METHOD PRIVATE PublishHmi
// Единый снимок состояния для внешней визуализации.
GVL_HMI.udiPlcHeartbeat := GVL_HMI.udiPlcHeartbeat + 1;
GVL_HMI.xHmiConnectionAlive := xHmiConnectionAlive;
GVL_HMI.xManualRecoveryActive := xManualRecoveryActive;
GVL_HMI.xGlobalError := GVL_CELL_CONTROL.xGlobalError;
GVL_HMI.xCellManual := GVL_CELL_CONTROL.xManual;
// Отказ тоже потребляет транзакцию: она не исполнится позже сама собой.
GVL_HMI.udiCellModeAckSeq := udiCellModeCommandSnapshot;
GVL_HMI.xErrorSimulationEnabled := GVL_CELL_SETTINGS.xErrorSimulationEnabled;
GVL_HMI.stSafetyFaultStatus := CELL_SAFETY.FaultStatus;
GVL_HMI.xSimulationAccelerationActive := GVL_CELL_SETTINGS.xSimulationAccelerationActive;
GVL_HMI.xSimulationAccelerationChangeAllowed := GVL_CELL_SETTINGS.xSimulationAccelerationChangeAllowed;
GVL_HMI.uiSimulationTimeFactorApplied := GVL_CELL_SETTINGS.uiSimulationTimeFactorApplied;
GVL_HMI.xSimulationAccelerationPending := GVL_CELL_SETTINGS.xSimulationAccelerationPending;
GVL_HMI.xSimulationAccelerationBusy := GVL_CELL_SETTINGS.xSimulationAccelerationBusy;
GVL_HMI.xSimulationAccelerationError := GVL_CELL_SETTINGS.xSimulationAccelerationError;
GVL_HMI.udiSimulationAccelerationErrorId := GVL_CELL_SETTINGS.udiSimulationAccelerationErrorId;
GVL_HMI.lrSafetyHomeX := GVL_POINT.Points[E_POINT_NAME.HOME_SAFETY].X;
GVL_HMI.lrSafetyHomeY := GVL_POINT.Points[E_POINT_NAME.HOME_SAFETY].Y;
GVL_HMI.lrSafetyHomeZ := GVL_POINT.Points[E_POINT_NAME.HOME_SAFETY].Z;
GVL_HMI.lrSafetyHomeSpeedFactor := GVL_POINT.Points[E_POINT_NAME.HOME_SAFETY].SpeedFactor;
GVL_HMI.lrSafetyHomeToleranceX := GVL_CELL_SETTINGS.lrSafetyHomeToleranceX;
GVL_HMI.lrSafetyHomeToleranceY := GVL_CELL_SETTINGS.lrSafetyHomeToleranceY;
GVL_HMI.lrSafetyHomeToleranceZ := GVL_CELL_SETTINGS.lrSafetyHomeToleranceZ;
GVL_HMI.rRobotAccelerationPercent := GVL_CELL_SETTINGS.rRobotAccelerationPercent;
GVL_HMI.rRobotDecelerationPercent := GVL_CELL_SETTINGS.rRobotDecelerationPercent;
GVL_HMI.rRobotJerkPercent := GVL_CELL_SETTINGS.rRobotJerkPercent;
GVL_HMI.lrRobotHaltDeceleration := GVL_CELL_SETTINGS.lrRobotHaltDeceleration;
GVL_HMI.lrRobotHaltJerk := GVL_CELL_SETTINGS.lrRobotHaltJerk;
GVL_HMI.stCellMachineTimeouts := GVL_CELL_SETTINGS.stMachineTimeouts;
GVL_HMI.stCellAxisTimeouts := GVL_CELL_SETTINGS.stAxisTimeouts;
GVL_HMI.stCellAxisGroupTimeouts := GVL_CELL_SETTINGS.stAxisGroupTimeouts;
GVL_HMI.tPointCheckStartTimeout := GVL_CELL_SETTINGS.tPointCheckStartTimeout;
GVL_HMI.tSimulationDynamicsTimeout := GVL_CELL_SETTINGS.tSimulationDynamicsTimeout;
GVL_HMI.tHmiWatchdogTimeout := GVL_CELL_SETTINGS.tHmiWatchdogTimeout;
GVL_HMI.tMobileMotionWatchdogTimeout := GVL_CELL_SETTINGS.tMobileMotionWatchdogTimeout;
GVL_HMI.tPointCheckWatchdogTimeout := GVL_CELL_SETTINGS.tPointCheckWatchdogTimeout;
GVL_HMI.tHmiCommandFreshnessTimeout := GVL_CELL_SETTINGS.tHmiCommandFreshnessTimeout;
GVL_HMI.tAlarmHornDuration := GVL_CELL_SETTINGS.tAlarmHornDuration;
GVL_HMI.tInputFilterRise := GVL_CELL_SETTINGS.tInputFilterRise;
GVL_HMI.tInputFilterFall := GVL_CELL_SETTINGS.tInputFilterFall;
GVL_HMI.xIoFilterSettingsChangeAllowed := GVL_CELL_SETTINGS.xIoFilterSettingsChangeAllowed;
GVL_HMI.xPhysicalIoActive := GVL_PHYSICAL_IO.xNormalActive
	AND (GVL_CELL_SETTINGS.eTestEnvironment = E_CELL_TEST_ENVIRONMENT.NORMAL);
GVL_HMI.xPhysicalIoMappingVerified := GVL_PHYSICAL_IO.xMappingVerified;
GVL_HMI.xCellSettingsChangeAllowed := GVL_CELL_SETTINGS.xCellSettingsChangeAllowed;
GVL_HMI.rPointCheckSpeedPercent := GVL_CELL_SETTINGS.rPointCheckSpeedPercent;
GVL_HMI.xPointCheckActive := xPointCheckActive;
IF xPointCheckActive THEN
	GVL_HMI.rPointCheckAppliedSpeedPercent := rPointCheckLatchedSpeed;
ELSE
	GVL_HMI.rPointCheckAppliedSpeedPercent := GVL_CELL_SETTINGS.rPointCheckSpeedPercent;
END_IF;
GVL_HMI.xPointTableReady := xPointTableReady;
GVL_HMI.astPointEditorPoints[1] := GVL_POINT.Points[E_POINT_NAME.MACHINE_1_ABOVE];
GVL_HMI.astPointEditorPoints[2] := GVL_POINT.Points[E_POINT_NAME.MACHINE_1_CHUCK_APROACH];
GVL_HMI.astPointEditorPoints[3] := GVL_POINT.Points[E_POINT_NAME.MACHINE_1_CHUCK_POSITION];
GVL_HMI.astPointEditorPoints[4] := GVL_POINT.Points[E_POINT_NAME.MACHINE_2_ABOVE];
GVL_HMI.astPointEditorPoints[5] := GVL_POINT.Points[E_POINT_NAME.MACHINE_2_CHUCK_APROACH];
GVL_HMI.astPointEditorPoints[6] := GVL_POINT.Points[E_POINT_NAME.MACHINE_2_CHUCK_POSITION];
GVL_HMI.astPointEditorPoints[7] := GVL_POINT.Points[E_POINT_NAME.MACHINE_3_ABOVE];
GVL_HMI.astPointEditorPoints[8] := GVL_POINT.Points[E_POINT_NAME.MACHINE_3_CHUCK_APROACH];
GVL_HMI.astPointEditorPoints[9] := GVL_POINT.Points[E_POINT_NAME.MACHINE_3_CHUCK_POSITION];
GVL_HMI.astPointEditorPoints[10] := GVL_POINT.Points[E_POINT_NAME.HOME_SAFETY];
GVL_HMI.astPointEditorPoints[11] := GVL_POINT.Points[E_POINT_NAME.MAGAZINE_1_DETAIL];
GVL_HMI.astPointEditorPoints[12] := GVL_POINT.Points[E_POINT_NAME.MAGAZINE_2_DETAIL];
GVL_HMI.astPointEditorPoints[13] := GVL_POINT.Points[E_POINT_NAME.GEOMETRY_1_PLACE];
GVL_HMI.astPointEditorPoints[14] := GVL_POINT.Points[E_POINT_NAME.GEOMETRY_2_PLACE];
GVL_HMI.auiPointEditorPointId[1] := TO_UINT(E_POINT_NAME.MACHINE_1_ABOVE);
GVL_HMI.auiPointEditorPointId[2] := TO_UINT(E_POINT_NAME.MACHINE_1_CHUCK_APROACH);
GVL_HMI.auiPointEditorPointId[3] := TO_UINT(E_POINT_NAME.MACHINE_1_CHUCK_POSITION);
GVL_HMI.auiPointEditorPointId[4] := TO_UINT(E_POINT_NAME.MACHINE_2_ABOVE);
GVL_HMI.auiPointEditorPointId[5] := TO_UINT(E_POINT_NAME.MACHINE_2_CHUCK_APROACH);
GVL_HMI.auiPointEditorPointId[6] := TO_UINT(E_POINT_NAME.MACHINE_2_CHUCK_POSITION);
GVL_HMI.auiPointEditorPointId[7] := TO_UINT(E_POINT_NAME.MACHINE_3_ABOVE);
GVL_HMI.auiPointEditorPointId[8] := TO_UINT(E_POINT_NAME.MACHINE_3_CHUCK_APROACH);
GVL_HMI.auiPointEditorPointId[9] := TO_UINT(E_POINT_NAME.MACHINE_3_CHUCK_POSITION);
GVL_HMI.auiPointEditorPointId[10] := TO_UINT(E_POINT_NAME.HOME_SAFETY);
GVL_HMI.auiPointEditorPointId[11] := TO_UINT(E_POINT_NAME.MAGAZINE_1_DETAIL);
GVL_HMI.auiPointEditorPointId[12] := TO_UINT(E_POINT_NAME.MAGAZINE_2_DETAIL);
GVL_HMI.auiPointEditorPointId[13] := TO_UINT(E_POINT_NAME.GEOMETRY_1_PLACE);
GVL_HMI.auiPointEditorPointId[14] := TO_UINT(E_POINT_NAME.GEOMETRY_2_PLACE);
GVL_HMI.xModbusMode := GVL_ROBOT_MODBUS.xModeActive;
GVL_HMI.xRobotModeChangeAllowed := GVL_ROBOT_MODBUS.xRobotModeChangeAllowed;
GVL_HMI.xModbusSettingsChangeAllowed := GVL_ROBOT_MODBUS.xSettingsChangeAllowed;
GVL_HMI.stRobotModbusStatus := GVL_ROBOT_MODBUS.Status;
uiMagazine := GVL_CELL_MANAGER.Status.uiActiveMagazine;
IF (uiMagazine < UINT#1) OR (uiMagazine > UINT#2) THEN
	uiMagazine := UINT#1;
END_IF;
GVL_HMI.stTestObservability.udiAppliedScenarioSeq := GVL_HMI.udiTestScenarioAckSeq;
GVL_HMI.stTestObservability.uiCellState := TO_UINT(GVL_CELL_MANAGER.Diag.eState);
GVL_HMI.stTestObservability.uiRobotState := TO_UINT(GVL_ROBOT.Diag.eState);
GVL_HMI.stTestObservability.uiRobotAction := TO_UINT(GVL_ROBOT.Diag.eActiveAction);
GVL_HMI.stTestObservability.uiRobotPoint := TO_UINT(GVL_ROBOT.Diag.eActivePoint);
GVL_HMI.stTestObservability.uiActiveMagazine := GVL_CELL_MANAGER.Status.uiActiveMagazine;
GVL_HMI.stTestObservability.uiMagazineState := TO_UINT(GVL_MAGAZINE.astDiag[uiMagazine].eState);
GVL_HMI.stTestObservability.uiMagazineOperation := TO_UINT(GVL_MAGAZINE.astStatus[uiMagazine].eActualOperation);
GVL_HMI.stTestObservability.uiTakeSlot := SINT_TO_UINT(GVL_MAGAZINE.astStatus[uiMagazine].iSelectedBlank);
GVL_HMI.stTestObservability.uiPutSlot := SINT_TO_UINT(GVL_MAGAZINE.astStatus[uiMagazine].iSelectedFreeSlot);
GVL_HMI.stTestObservability.uiSelectedMachine := GVL_CELL_MANAGER.Status.uiSelectedMachine;
GVL_HMI.stTestObservability.uiSelectedType := GVL_MULTI_TYPE.CycleStatus.uiSelectedType;
GVL_HMI.stTestObservability.uiErrorSource := UINT#0;
GVL_HMI.stTestObservability.dwErrorCode := DWORD#0;
FOR uiMachine := 1 TO 3 DO
	GVL_HMI.stTestObservability.auiMachineState[uiMachine] := TO_UINT(GVL_MACHINE.Diag[uiMachine].eState);
	GVL_HMI.stTestObservability.auiMachineOperation[uiMachine] := TO_UINT(GVL_MACHINE.Diag[uiMachine].eActualOperation);
END_FOR;
IF GVL_ROBOT.Error.dwErrorActive <> DWORD#0 THEN
	GVL_HMI.stTestObservability.uiErrorSource := UINT#2;
	GVL_HMI.stTestObservability.dwErrorCode := GVL_ROBOT.Error.dwErrorActive;
ELSIF GVL_MAGAZINE.astError[1].dwErrorActive <> DWORD#0 THEN
	GVL_HMI.stTestObservability.uiErrorSource := UINT#3;
GVL_HMI.stTestObservability.dwErrorCode := GVL_MAGAZINE.astError[1].dwErrorActive;
ELSIF GVL_MAGAZINE.astError[2].dwErrorActive <> DWORD#0 THEN
	GVL_HMI.stTestObservability.uiErrorSource := UINT#7;
	GVL_HMI.stTestObservability.dwErrorCode := GVL_MAGAZINE.astError[2].dwErrorActive;
ELSIF GVL_CELL_MANAGER.Error.dwErrorActive <> DWORD#0 THEN
	GVL_HMI.stTestObservability.uiErrorSource := UINT#1;
	GVL_HMI.stTestObservability.dwErrorCode := GVL_CELL_MANAGER.Error.dwErrorActive;
ELSE
	FOR uiMachine := 1 TO 3 DO
		IF GVL_MACHINE.Error[uiMachine].dwErrorActive <> DWORD#0 THEN
			GVL_HMI.stTestObservability.uiErrorSource := uiMachine + UINT#3;
			GVL_HMI.stTestObservability.dwErrorCode := GVL_MACHINE.Error[uiMachine].dwErrorActive;
		END_IF;
	END_FOR;
END_IF;
FOR uiMachine := 1 TO 9 DO
	GVL_HMI.auiRobotModbusWriteRegisters[uiMachine] :=
		GVL_ROBOT_MODBUS.auiWriteRegisters[uiMachine - 1];
END_FOR;
FOR uiMachine := 1 TO 17 DO
	GVL_HMI.auiRobotModbusReadRegisters[uiMachine] :=
		GVL_ROBOT_MODBUS.auiReadRegisters[uiMachine - 1];
END_FOR;
GVL_HMI.xSimAxisGroupErrorAllowed := GVL_AXIS_GROUP.AxisGroup.Status.xSimErrorAllowed;
GVL_HMI.astAxisFaultStatus[1] := AXIS_X.FaultStatus;
GVL_HMI.astAxisFaultStatus[2] := AXIS_Y.FaultStatus;
GVL_HMI.astAxisFaultStatus[3] := AXIS_Z.FaultStatus;
GVL_HMI.stAxisGroupFaultStatus := GROUP_XYZ.FaultStatus;
GVL_HMI.stGripperFaultStatus := ROBOT.FaultStatus.stGripper;
GVL_HMI.stRobotFaultStatus := ROBOT.FaultStatus.stRobot;
GVL_HMI.stCellFaultStatus := CELL_MANAGER.FaultStatus;
GVL_HMI.stPointFaultStatus := ROBOT.FaultStatus.stPoint;
GVL_HMI.stMagazineFaultStatus := fbMagazine1.FaultStatus;
GVL_HMI.astMagazineFaultStatus[1] := fbMagazine1.FaultStatus;
GVL_HMI.astMagazineFaultStatus[2] := fbMagazine2.FaultStatus;
GVL_HMI.rLoadCNC_1 := GVL_STATISTIC.stStatistic.stMachineStat.rLoadCNC_1;
GVL_HMI.rLoadCNC_2 := GVL_STATISTIC.stStatistic.stMachineStat.rLoadCNC_2;
GVL_HMI.rLoadCNC_3 := GVL_STATISTIC.stStatistic.stMachineStat.rLoadCNC_3;
GVL_HMI.rRobot := GVL_STATISTIC.stStatistic.stRobotStat.rRobot;

GVL_HMI.stCellStatus := GVL_CELL_MANAGER.Status;
GVL_HMI.stCellStatus.xResetAllowed := xAlarmResetAllowed;
GVL_HMI.stCellDiag := GVL_CELL_MANAGER.Diag;
GVL_HMI.stCellError := GVL_CELL_MANAGER.Error;
GVL_HMI.stCellSafetyStatus := CELL_SAFETY.Status;
GVL_HMI.stCellSafetyDiag := CELL_SAFETY.Diag;
GVL_HMI.stCellSafetyError := CELL_SAFETY.Error;
GVL_HMI.astButtonStationIoStatus := CELL_SAFETY.astButtonStationIoStatus;
GVL_HMI.stFrontControlCabinetIoStatus := CELL_SAFETY.stFrontControlCabinetIoStatus;
GVL_HMI.xSignalTowerRed := GVL_CELL_SAFETY_IO.xSignalTowerRedOutput;
GVL_HMI.xSignalTowerAmber := GVL_CELL_SAFETY_IO.xSignalTowerAmberOutput;
GVL_HMI.xSignalTowerGreen := GVL_CELL_SAFETY_IO.xSignalTowerGreenOutput;
GVL_HMI.stRearControlCabinetIoStatus := CELL_SAFETY.stRearControlCabinetIoStatus;
GVL_HMI.stMpgIoStatus := CELL_SAFETY.stMpgIoStatus;
GVL_HMI.astEnclosureDoorStatus := CELL_SAFETY.astEnclosureDoorStatus;
GVL_HMI.stMultiType.Config := GVL_MULTI_TYPE.Config;
GVL_HMI.stMultiType.ConfigStatus := GVL_MULTI_TYPE.ConfigStatus;
GVL_HMI.stMultiType.CycleStatus := GVL_MULTI_TYPE.CycleStatus;

GVL_HMI.stRobotStatus := GVL_ROBOT.Status;
GVL_HMI.stRobotDiag := GVL_ROBOT.Diag;
GVL_HMI.stRobotError := GVL_ROBOT.Error;
GVL_HMI.stGripperDiag := GVL_ROBOT.GripperDiag;
GVL_HMI.stGripperError := GVL_ROBOT.GripperError;
GVL_HMI.stAxisGroupStatus := GVL_AXIS_GROUP.AxisGroup.Status;
GVL_HMI.stAxisGroupDiag := GVL_AXIS_GROUP.AxisGroup.Diag;
GVL_HMI.stAxisGroupError := GVL_AXIS_GROUP.AxisGroup.Error;
GVL_HMI.stMotionManagerStatus := GVL_MOTION_MANAGER.stMotionManager.Status;
GVL_HMI.stMotionManagerDiag := GVL_MOTION_MANAGER.stMotionManager.Diag;
GVL_HMI.stMotionManagerError := GVL_MOTION_MANAGER.stMotionManager.Error;
GVL_HMI.stPointManagerStatus := GVL_POINT_MANAGER.PointManager.Status;
GVL_HMI.stPointManagerDiag := GVL_POINT_MANAGER.PointManager.Diag;
GVL_HMI.stPointManagerError := GVL_POINT_MANAGER.PointManager.Error;

FOR uiMachine := 1 TO 3 DO
	GVL_HMI.astAxisStatus[uiMachine] := GVL_AXIS.arrAxis[uiMachine].Status;
	GVL_HMI.astAxisDiag[uiMachine] := GVL_AXIS.arrAxis[uiMachine].Diag;
	GVL_HMI.astAxisError[uiMachine] := GVL_AXIS.arrAxis[uiMachine].Error;
END_FOR;

GVL_HMI.stMagazineStatus := GVL_MAGAZINE.astStatus[1];
GVL_HMI.stMagazineDiag := GVL_MAGAZINE.astDiag[1];
GVL_HMI.stMagazineError := GVL_MAGAZINE.astError[1];
FOR uiMagazine := UINT#1 TO UINT#2 DO
	GVL_HMI.astMagazineStatus[uiMagazine] := GVL_MAGAZINE.astStatus[uiMagazine];
	GVL_HMI.astMagazineDiag[uiMagazine] := GVL_MAGAZINE.astDiag[uiMagazine];
	GVL_HMI.astMagazineError[uiMagazine] := GVL_MAGAZINE.astError[uiMagazine];
	GVL_HMI.astMagazineInventory[uiMagazine] := GVL_DETAIL.astMagazine[uiMagazine];
END_FOR;
GVL_HMI.stAlarmStatus := GVL_ALARM.Status;
GVL_HMI.astAlarmEvent := GVL_ALARM.Events;

FOR uiMachine := 1 TO 3 DO
	GVL_HMI.astMachineStatus[uiMachine] := GVL_MACHINE.Status[uiMachine];
	GVL_HMI.astMachineDiag[uiMachine] := GVL_MACHINE.Diag[uiMachine];
	GVL_HMI.astMachineError[uiMachine] := GVL_MACHINE.Error[uiMachine];
	CASE uiMachine OF
		1:
			GVL_HMI.astMachineFaultStatus[uiMachine] := MACHINE_1_FAULT.Status;
			GVL_HMI.astMachineFaultStatus[uiMachine].xResetAllowed :=
				MACHINE_1_SIM.Diag.xResetAllowed OR GVL_MACHINE.Status[uiMachine].xResetAllowed;
		2:
			GVL_HMI.astMachineFaultStatus[uiMachine] := MACHINE_2_FAULT.Status;
			GVL_HMI.astMachineFaultStatus[uiMachine].xResetAllowed :=
				MACHINE_2_SIM.Diag.xResetAllowed OR GVL_MACHINE.Status[uiMachine].xResetAllowed;
		3:
			GVL_HMI.astMachineFaultStatus[uiMachine] := MACHINE_3_FAULT.Status;
			GVL_HMI.astMachineFaultStatus[uiMachine].xResetAllowed :=
				MACHINE_3_SIM.Diag.xResetAllowed OR GVL_MACHINE.Status[uiMachine].xResetAllowed;
	END_CASE;
END_FOR;

GVL_HMI.astMachineIoStatus[1] := MACHINE_1_FAULT.MachineStatus;
GVL_HMI.astMachineIoStatus[2] := MACHINE_2_FAULT.MachineStatus;
GVL_HMI.astMachineIoStatus[3] := MACHINE_3_FAULT.MachineStatus;
GVL_HMI.astMachineRawIoStatus[1] := MACHINE_1_SIM.Status;
GVL_HMI.astMachineRawIoStatus[2] := MACHINE_2_SIM.Status;
GVL_HMI.astMachineRawIoStatus[3] := MACHINE_3_SIM.Status;
GVL_HMI.astMachineTimeouts[1] := MACHINE_1_FAULT.Timeouts;
GVL_HMI.astMachineTimeouts[2] := MACHINE_2_FAULT.Timeouts;
GVL_HMI.astMachineTimeouts[3] := MACHINE_3_FAULT.Timeouts;
GVL_HMI.astMachineSimDiag[1] := MACHINE_1_SIM.Diag;
GVL_HMI.astMachineSimDiag[2] := MACHINE_2_SIM.Diag;
GVL_HMI.astMachineSimDiag[3] := MACHINE_3_SIM.Diag;
GVL_HMI.astMachineSimError[1] := MACHINE_1_SIM.Error;
GVL_HMI.astMachineSimError[2] := MACHINE_2_SIM.Error;
GVL_HMI.astMachineSimError[3] := MACHINE_3_SIM.Error;

FOR iDetail := 1 TO GVL_CELL_SETTINGS.NumberDetail DO
	GVL_HMI.astMagazineSlot[iDetail] := GVL_DETAIL.astMagazine[1].aSlots[iDetail];
END_FOR;

// Ack only the snapshot actually dispatched through all consumers this scan.
FOR uiHmiCommandIndex := UINT#1 TO UINT#121 DO
	IF axHmiCommandConsumed[uiHmiCommandIndex] THEN
		GVL_HMI.audiHmiCommandAckSeq[uiHmiCommandIndex] := audiHmiCommandSnapshot[uiHmiCommandIndex];
	END_IF;
END_FOR;
GVL_HMI.udiCellSettingAckSeq := udiCellSettingSnapshot;

GVL_HMI.uiMagazineMode := GVL_TWO_PALLET.uiMode;
GVL_HMI.xMagazineModeAllowed := GVL_TWO_PALLET.xModeChangeAllowed;
GVL_HMI.astTwinStatus := GVL_TWO_PALLET.astStatus;
GVL_HMI.astTwinConfig := GVL_TWO_PALLET.astActiveConfig;
GVL_HMI.astTwinStore := GVL_TWO_PALLET.astStore;
END_METHOD

METHOD PRIVATE IsHmiCommandFresh : BOOL
VAR_INPUT
	udiIssuedAtMs : UDINT;
END_VAR
VAR
	uliAgeMs : ULINT;
END_VAR
// Explicit modulo-2^32 age: TIME() rolls over after about 49 days.
IF udiHmiCommandNowMs >= udiIssuedAtMs THEN
	uliAgeMs := UDINT_TO_ULINT(udiHmiCommandNowMs) - UDINT_TO_ULINT(udiIssuedAtMs);
ELSE
	uliAgeMs := ULINT#4294967296 + UDINT_TO_ULINT(udiHmiCommandNowMs) - UDINT_TO_ULINT(udiIssuedAtMs);
END_IF;
IsHmiCommandFresh := uliAgeMs <= UDINT_TO_ULINT(
	TIME_TO_UDINT(GVL_CELL_SETTINGS.tHmiCommandFreshnessTimeout)
);
END_METHOD

METHOD PRIVATE WritePhysicalOutputs
// Единственная страница назначения выходов. Выполняется после всех владельцев команд.
// Не публикуем команды симулятора на железо при смене среды в текущем скане.
xPhysicalOutputEnable := GVL_PHYSICAL_IO.xNormalActive
	AND (GVL_CELL_SETTINGS.eTestEnvironment = E_CELL_TEST_ENVIRONMENT.NORMAL);
IF xPhysicalOutputEnable THEN
	FOR uiMachine := 1 TO 3 DO
		IF GVL_MACHINE.Command[uiMachine].stIo.xCloseDoor
		AND NOT GVL_MACHINE.Command[uiMachine].stIo.xOpenDoor THEN
			GVL_PHYSICAL_IO.axMachineHatchClose[uiMachine] := TRUE;
		ELSIF GVL_MACHINE.Command[uiMachine].stIo.xOpenDoor
		AND NOT GVL_MACHINE.Command[uiMachine].stIo.xCloseDoor THEN
			GVL_PHYSICAL_IO.axMachineHatchClose[uiMachine] := FALSE;
		ELSIF NOT xPhysicalOutputWasEnabled THEN
			GVL_PHYSICAL_IO.axMachineHatchClose[uiMachine] := GVL_MACHINE.astPhysicalInput[uiMachine].xDoorClosed;
		END_IF;
	END_FOR;
	IF NOT GVL_HMI.xModbusMode AND GVL_PHYSICAL_IO.stGripperCommand.xExecute THEN
		CASE GVL_PHYSICAL_IO.stGripperCommand.eAction OF
			E_ROBOT_ACTION.UNCLAMP_1: axIoGripperBase[1] := TRUE;
			E_ROBOT_ACTION.CLAMP_1: axIoGripperBase[1] := FALSE;
			E_ROBOT_ACTION.UNCLAMP_2: axIoGripperBase[2] := TRUE;
			E_ROBOT_ACTION.CLAMP_2: axIoGripperBase[2] := FALSE;
			E_ROBOT_ACTION.ROTATE_TO_BLANK: axIoGripperBase[3] := FALSE;
			E_ROBOT_ACTION.ROTATE_TO_DETAIL: axIoGripperBase[3] := TRUE;
		END_CASE;
	END_IF;
END_IF;
// Внешний SC-500 остаётся единственным владельцем захватов в Modbus.
IF NOT xPhysicalOutputEnable OR GVL_HMI.xModbusMode THEN
	axIoGripperBase[1] := FALSE;
	axIoGripperBase[2] := FALSE;
	axIoGripperBase[3] := FALSE;
END_IF;
GVL_PHYSICAL_IO.xDoGripper1Open := axIoGripperBase[1];
GVL_PHYSICAL_IO.xDoGripper2Open := axIoGripperBase[2];
GVL_PHYSICAL_IO.xDoRotateToDetail := axIoGripperBase[3];

GVL_PHYSICAL_IO.xDoMachine1HatchClosed := xPhysicalOutputEnable AND GVL_PHYSICAL_IO.axMachineHatchClose[1];
GVL_PHYSICAL_IO.xDoMachine1HatchUnLock := xPhysicalOutputEnable AND GVL_MACHINE.Command[1].stIo.xHatchUnLock;
GVL_PHYSICAL_IO.xDoMachine1ClampChuck := xPhysicalOutputEnable AND GVL_MACHINE.Command[1].stIo.xClampChuck AND NOT GVL_MACHINE.Command[1].stIo.xUnclampChuck;
GVL_PHYSICAL_IO.xDoMachine1UnclampChuck := xPhysicalOutputEnable AND GVL_MACHINE.Command[1].stIo.xUnclampChuck AND NOT GVL_MACHINE.Command[1].stIo.xClampChuck;
GVL_PHYSICAL_IO.xDoMachine1StartCycle := xPhysicalOutputEnable AND GVL_MACHINE.Command[1].stIo.xStartCycle;
GVL_PHYSICAL_IO.xDoMachine2HatchClosed := xPhysicalOutputEnable AND GVL_PHYSICAL_IO.axMachineHatchClose[2];
GVL_PHYSICAL_IO.xDoMachine2HatchUnLock := xPhysicalOutputEnable AND GVL_MACHINE.Command[2].stIo.xHatchUnLock;
GVL_PHYSICAL_IO.xDoMachine2ClampChuck := xPhysicalOutputEnable AND GVL_MACHINE.Command[2].stIo.xClampChuck AND NOT GVL_MACHINE.Command[2].stIo.xUnclampChuck;
GVL_PHYSICAL_IO.xDoMachine2UnclampChuck := xPhysicalOutputEnable AND GVL_MACHINE.Command[2].stIo.xUnclampChuck AND NOT GVL_MACHINE.Command[2].stIo.xClampChuck;
GVL_PHYSICAL_IO.xDoMachine2StartCycle := xPhysicalOutputEnable AND GVL_MACHINE.Command[2].stIo.xStartCycle;
GVL_PHYSICAL_IO.xDoMachine3HatchClosed := xPhysicalOutputEnable AND GVL_PHYSICAL_IO.axMachineHatchClose[3];
GVL_PHYSICAL_IO.xDoMachine3HatchUnLock := xPhysicalOutputEnable AND GVL_MACHINE.Command[3].stIo.xHatchUnLock;
GVL_PHYSICAL_IO.xDoMachine3ClampChuck := xPhysicalOutputEnable AND GVL_MACHINE.Command[3].stIo.xClampChuck AND NOT GVL_MACHINE.Command[3].stIo.xUnclampChuck;
GVL_PHYSICAL_IO.xDoMachine3UnclampChuck := xPhysicalOutputEnable AND GVL_MACHINE.Command[3].stIo.xUnclampChuck AND NOT GVL_MACHINE.Command[3].stIo.xClampChuck;
GVL_PHYSICAL_IO.xDoMachine3StartCycle := xPhysicalOutputEnable AND GVL_MACHINE.Command[3].stIo.xStartCycle;
GVL_PHYSICAL_IO.xDoDoor1Unlock := xPhysicalOutputEnable AND GVL_CELL_SAFETY_IO.axDoorUnlockOutput[1];
GVL_PHYSICAL_IO.xDoDoor2Unlock := xPhysicalOutputEnable AND GVL_CELL_SAFETY_IO.axDoorUnlockOutput[2];
GVL_PHYSICAL_IO.xDoDoor3Unlock := xPhysicalOutputEnable AND GVL_CELL_SAFETY_IO.axDoorUnlockOutput[3];
GVL_PHYSICAL_IO.xDoDoor4Unlock := xPhysicalOutputEnable AND GVL_CELL_SAFETY_IO.axDoorUnlockOutput[4];
GVL_PHYSICAL_IO.xDoSafetyRelayReset := xPhysicalOutputEnable AND GVL_CELL_SAFETY_IO.xSafetyRelayResetOutput;
GVL_PHYSICAL_IO.xDoSignalTowerGreenOutput := xPhysicalOutputEnable AND GVL_CELL_SAFETY_IO.xSignalTowerGreenOutput;
GVL_PHYSICAL_IO.xDoSignalTowerAmberOutput := xPhysicalOutputEnable AND GVL_CELL_SAFETY_IO.xSignalTowerAmberOutput;
GVL_PHYSICAL_IO.xDoSignalTowerRedOutput := xPhysicalOutputEnable AND GVL_CELL_SAFETY_IO.xSignalTowerRedOutput;
GVL_PHYSICAL_IO.xDoDoor1ButtonLamp := xPhysicalOutputEnable AND GVL_CELL_SAFETY_IO.axDoorButtonLampOutput[1];
GVL_PHYSICAL_IO.xDoDoor2ButtonLamp := xPhysicalOutputEnable AND GVL_CELL_SAFETY_IO.axDoorButtonLampOutput[2];
GVL_PHYSICAL_IO.xDoDoor3ButtonLamp := xPhysicalOutputEnable AND GVL_CELL_SAFETY_IO.axDoorButtonLampOutput[3];
GVL_PHYSICAL_IO.xDoDoor4ButtonLamp := xPhysicalOutputEnable AND GVL_CELL_SAFETY_IO.axDoorButtonLampOutput[4];
GVL_PHYSICAL_IO.xDoMagazine1LockIn := xPhysicalOutputEnable AND (GVL_TWO_PALLET.uiMode = UINT#1) AND GVL_TWO_PALLET.astOutput[1].xLockIn AND NOT GVL_TWO_PALLET.astOutput[1].xLockOut;
GVL_PHYSICAL_IO.xDoMagazine1LockOut := xPhysicalOutputEnable AND (GVL_TWO_PALLET.uiMode = UINT#1) AND GVL_TWO_PALLET.astOutput[1].xLockOut AND NOT GVL_TWO_PALLET.astOutput[1].xLockIn;
GVL_PHYSICAL_IO.xDoMagazine1StopIn := xPhysicalOutputEnable AND (GVL_TWO_PALLET.uiMode = UINT#1) AND GVL_TWO_PALLET.astOutput[1].xStopIn AND NOT GVL_TWO_PALLET.astOutput[1].xStopOut;
GVL_PHYSICAL_IO.xDoMagazine1StopOut := xPhysicalOutputEnable AND (GVL_TWO_PALLET.uiMode = UINT#1) AND GVL_TWO_PALLET.astOutput[1].xStopOut AND NOT GVL_TWO_PALLET.astOutput[1].xStopIn;
GVL_PHYSICAL_IO.xDoMagazine1LiftUp := xPhysicalOutputEnable AND (GVL_TWO_PALLET.uiMode = UINT#1) AND GVL_TWO_PALLET.astOutput[1].xLiftUp AND NOT GVL_TWO_PALLET.astOutput[1].xLiftDown;
GVL_PHYSICAL_IO.xDoMagazine1LiftDown := xPhysicalOutputEnable AND (GVL_TWO_PALLET.uiMode = UINT#1) AND GVL_TWO_PALLET.astOutput[1].xLiftDown AND NOT GVL_TWO_PALLET.astOutput[1].xLiftUp;
GVL_PHYSICAL_IO.xDoMagazine2LockIn := xPhysicalOutputEnable AND (GVL_TWO_PALLET.uiMode = UINT#1) AND GVL_TWO_PALLET.astOutput[2].xLockIn AND NOT GVL_TWO_PALLET.astOutput[2].xLockOut;
GVL_PHYSICAL_IO.xDoMagazine2LockOut := xPhysicalOutputEnable AND (GVL_TWO_PALLET.uiMode = UINT#1) AND GVL_TWO_PALLET.astOutput[2].xLockOut AND NOT GVL_TWO_PALLET.astOutput[2].xLockIn;
GVL_PHYSICAL_IO.xDoMagazine2StopIn := xPhysicalOutputEnable AND (GVL_TWO_PALLET.uiMode = UINT#1) AND GVL_TWO_PALLET.astOutput[2].xStopIn AND NOT GVL_TWO_PALLET.astOutput[2].xStopOut;
GVL_PHYSICAL_IO.xDoMagazine2StopOut := xPhysicalOutputEnable AND (GVL_TWO_PALLET.uiMode = UINT#1) AND GVL_TWO_PALLET.astOutput[2].xStopOut AND NOT GVL_TWO_PALLET.astOutput[2].xStopIn;
GVL_PHYSICAL_IO.xDoMagazine2LiftUp := xPhysicalOutputEnable AND (GVL_TWO_PALLET.uiMode = UINT#1) AND GVL_TWO_PALLET.astOutput[2].xLiftUp AND NOT GVL_TWO_PALLET.astOutput[2].xLiftDown;
GVL_PHYSICAL_IO.xDoMagazine2LiftDown := xPhysicalOutputEnable AND (GVL_TWO_PALLET.uiMode = UINT#1) AND GVL_TWO_PALLET.astOutput[2].xLiftDown AND NOT GVL_TWO_PALLET.astOutput[2].xLiftUp;


GVL_PHYSICAL_IO.xDoCellAlarmHorn := xPhysicalOutputEnable AND GVL_CELL_SAFETY_IO.xAlarmHornOutput;
GVL_PHYSICAL_IO.xDoGk1DriveRun := xPhysicalOutputEnable AND GEOMETRY[1].xRunOutput;
GVL_PHYSICAL_IO.xDoGk1DriveReset := xPhysicalOutputEnable AND GEOMETRY[1].xResetOutput;

GVL_PHYSICAL_IO.xDoGk2DriveRun := xPhysicalOutputEnable AND GEOMETRY[2].xRunOutput;
GVL_PHYSICAL_IO.xDoGk2DriveReset := xPhysicalOutputEnable AND GEOMETRY[2].xResetOutput;

ApplyIoOutputOverrides();

xPhysicalOutputWasEnabled := xPhysicalOutputEnable;
END_METHOD

END_PROGRAM

// Device/Application/FB/FB_GEOMETRY_CONTROL
FUNCTION_BLOCK FB_GEOMETRY_CONTROL
VAR_INPUT
	xInitialize : BOOL;
	uiAction : UINT;
	xSupported : BOOL;
	xSimulation : BOOL;
	xGlobalError : BOOL;
	xManual : BOOL;
	xCellRunning : BOOL;
	xRobotBusy : BOOL;
	xMotionBusy : BOOL;
	xHmiAlive : BOOL;
	xIoManual : BOOL;
	xReset : BOOL;
	xDriveAlarm : BOOL;
	xDriveRunning : BOOL;
	xPartAtEnd : BOOL;
	rSimulationTravel : REAL;
	Signals : ST_GEOMETRY_SIGNALS;
	Config : ST_GEOMETRY_CONFIG;
	tTransport : TIME;
	tFeedback : TIME;
	tResetPulse : TIME;
	uiTimeFactor : UINT := UINT#1;
END_VAR
VAR_IN_OUT
	Memory : ST_GEOMETRY_MEMORY;
END_VAR
VAR_OUTPUT
	Status : ST_GEOMETRY_STATUS;
	Warning : ST_WARNING_EVENT;
	xRunOutput : BOOL;
	xResetOutput : BOOL;
	xCommandAccepted : BOOL;
	xSimulationEmptyConfirmed : BOOL; // Одноцикловое принятое изъятие/подтверждение пустоты виртуальной ленты
END_VAR
VAR
	xInitialized : BOOL;
	xEnabled : BOOL;
	xReserved : BOOL;
	xTransport : BOOL;
	xManualRun : BOOL;
	xDisablePending : BOOL;
	xEnableWanted : BOOL;
	xResetBusy : BOOL;
	xResetSeen : BOOL;
	xConfigurationValid : BOOL;
	xManualBase : BOOL;
	xCommandRejected : BOOL;
	dwControlBlockers : DWORD;
	tTransportScaled : TIME;
	tFeedbackScaled : TIME;
	tonTransport : TON;
	tonFeedback : TON;
	tonRemoved : TON;
	tonReset : TON;
	stRemoved : ST_GEOMETRY_CALL;
END_VAR

IF xInitialize THEN xInitialized := FALSE; END_IF;
IF NOT xInitialized THEN
	// После рестарта конечный датчик не доказывает пустоту всей ленты.
	xEnabled := FALSE; xReserved := FALSE; xTransport := FALSE; xManualRun := FALSE;
	xDisablePending := FALSE; xEnableWanted := FALSE; xResetBusy := FALSE; xResetSeen := FALSE;
	Memory.xRecoveryRequired := TRUE; xInitialized := TRUE;
END_IF;
xCommandAccepted := FALSE;
xSimulationEmptyConfirmed := FALSE;
xCommandRejected := FALSE;
xConfigurationValid := Config.xConfigured AND (Config.lrSpeedFactor >= 0.1)
	AND (Config.lrSpeedFactor <= 1.0) AND (Config.lrSafeZ < 0.0) AND (Config.lrSafeZ >= -10000.0);
tTransportScaled := UDINT_TO_TIME(MAX(UDINT#1, TIME_TO_UDINT(tTransport) / UINT_TO_UDINT(MAX(UINT#1, uiTimeFactor))));
tFeedbackScaled := UDINT_TO_TIME(MAX(UDINT#1, TIME_TO_UDINT(tFeedback) / UINT_TO_UDINT(MAX(UINT#1, uiTimeFactor))));

IF xDriveAlarm THEN Memory.dwAlarm := Memory.dwAlarm OR DWORD#1; END_IF;
IF Memory.dwAlarm <> DWORD#0 THEN
	Memory.xRecoveryRequired := TRUE;
	IF Signals.xRobotInteraction THEN Memory.xRobotStopLatched := TRUE; END_IF;
	xEnabled := FALSE; xEnableWanted := FALSE; xTransport := FALSE; xManualRun := FALSE;
END_IF;
IF xGlobalError OR NOT xSupported OR xIoManual THEN
	IF Memory.xOccupied OR xReserved OR xTransport OR xManualRun THEN Memory.xRecoveryRequired := TRUE; END_IF;
	xEnabled := FALSE; xEnableWanted := FALSE; xTransport := FALSE; xManualRun := FALSE;
	xResetBusy := FALSE;
END_IF;
IF NOT xHmiAlive OR NOT xManual OR xCellRunning THEN xManualRun := FALSE; END_IF;

IF Signals.xReserve AND xEnabled AND xConfigurationValid AND NOT Memory.xOccupied
	AND NOT Memory.xRecoveryRequired AND NOT xPartAtEnd AND NOT xDriveRunning
	AND NOT xManualRun AND NOT xResetBusy AND NOT xGlobalError AND xSupported AND NOT xIoManual
	AND (Memory.dwAlarm = DWORD#0) THEN
	xReserved := TRUE; Memory.Part := Signals.Call;
END_IF;
IF Signals.xDeposited AND xReserved AND (Signals.Call.udiId <> UDINT#0)
	AND (Memory.udiLastDepositId <> Signals.Call.udiId) THEN
	Memory.xOccupied := TRUE; Memory.xAtEndSeen := FALSE;
	Memory.udiLastDepositId := Signals.Call.udiId;
	Memory.udiProducedPartsTotal := Memory.udiProducedPartsTotal + UDINT#1;
	Memory.Part := Signals.Call; Memory.Part.uiState := UINT#4;
	IF (Memory.Part.uiMachine >= UINT#1) AND (Memory.Part.uiMachine <= UINT#3) THEN
		GVL_GEOMETRY_CONTROL.astCalls[Memory.Part.uiMachine] := Memory.Part;
	END_IF;
	F_GEOMETRY_EVENT(Call := Memory.Part);
END_IF;
IF Signals.xReleased THEN
	xReserved := FALSE;
	IF Memory.xOccupied AND xEnabled AND NOT xDisablePending AND NOT Memory.xRecoveryRequired
		AND (Memory.dwAlarm = DWORD#0) AND NOT xGlobalError THEN xTransport := TRUE; END_IF;
END_IF;

xManualBase := xSupported AND xManual AND NOT xCellRunning AND NOT xRobotBusy
	AND NOT xMotionBusy AND NOT Signals.xRobotInteraction AND NOT xReserved
	AND xHmiAlive AND NOT xGlobalError AND NOT xIoManual AND NOT xResetBusy;
Status.xConfigAllowed := xManualBase AND NOT xEnabled AND NOT xDriveRunning AND NOT Memory.xOccupied;
// Допуск записи данных публикует RunGeometryControl независимо от состояния ГК.
// xConfigAllowed остаётся строгим допуском проверки с движением к базе.
// Включение и подтверждение пустоты зависят от выбранного ГК.
// Движение робота вне этой станции и работа ячейки не запрещают эти команды.
// Биты причин в astGeometryStatus: контракт описан в DOKS/24-geometry-control.md.
dwControlBlockers := DWORD#0;
IF NOT xSupported THEN dwControlBlockers := dwControlBlockers OR DWORD#1; END_IF;
IF NOT xHmiAlive THEN dwControlBlockers := dwControlBlockers OR DWORD#2; END_IF;
IF xGlobalError THEN dwControlBlockers := dwControlBlockers OR DWORD#4; END_IF;
IF xIoManual THEN dwControlBlockers := dwControlBlockers OR DWORD#8; END_IF;
IF Memory.dwAlarm <> DWORD#0 THEN dwControlBlockers := dwControlBlockers OR DWORD#16; END_IF;
IF Signals.xRobotInteraction THEN dwControlBlockers := dwControlBlockers OR DWORD#64; END_IF;
IF xReserved THEN dwControlBlockers := dwControlBlockers OR DWORD#128; END_IF;
IF xDriveRunning THEN dwControlBlockers := dwControlBlockers OR DWORD#256; END_IF;
IF xManualRun THEN dwControlBlockers := dwControlBlockers OR DWORD#512; END_IF;
IF xResetBusy THEN dwControlBlockers := dwControlBlockers OR DWORD#1024; END_IF;
IF xDisablePending THEN dwControlBlockers := dwControlBlockers OR DWORD#2048; END_IF;
IF xTransport THEN dwControlBlockers := dwControlBlockers OR DWORD#8192; END_IF;
Status.dwEnableBlockers := dwControlBlockers;
IF NOT xConfigurationValid THEN Status.dwEnableBlockers := Status.dwEnableBlockers OR DWORD#32; END_IF;
IF xEnabled THEN Status.dwEnableBlockers := Status.dwEnableBlockers OR DWORD#4096; END_IF;
Status.xEnableAllowed := Status.dwEnableBlockers = DWORD#0;
Status.xDisableAllowed := xSupported AND (xEnabled OR xEnableWanted OR xDisablePending);
Status.dwConfirmBlockers := dwControlBlockers;
IF xEnableWanted AND NOT xConfigurationValid THEN Status.dwConfirmBlockers := Status.dwConfirmBlockers OR DWORD#32; END_IF;
IF NOT xEnableWanted AND NOT Memory.xRecoveryRequired THEN Status.dwConfirmBlockers := Status.dwConfirmBlockers OR DWORD#16384; END_IF;
IF xPartAtEnd THEN Status.dwConfirmBlockers := Status.dwConfirmBlockers OR DWORD#32768; END_IF;
Status.xConfirmAllowed := Status.dwConfirmBlockers = DWORD#0;
Status.xManualStartAllowed := xManualBase AND NOT xDriveAlarm AND (Memory.dwAlarm = DWORD#0) AND NOT xManualRun;
Status.xResetAllowed := (Memory.dwAlarm <> DWORD#0) AND NOT xResetBusy AND xSupported
	AND NOT xGlobalError AND NOT xIoManual
	AND NOT xRobotBusy AND NOT xMotionBusy AND NOT xManualRun AND NOT xTransport;
Status.xSimulationRemoveAllowed := xSimulation AND xSupported AND xHmiAlive
	AND NOT xGlobalError AND NOT xIoManual AND NOT xResetBusy
	AND Memory.xOccupied AND NOT Signals.xRobotInteraction AND NOT xReserved AND NOT xDriveRunning;

CASE uiAction OF
	UINT#1:
		IF Status.xEnableAllowed THEN
			IF Memory.xRecoveryRequired OR Memory.xOccupied OR xPartAtEnd THEN
				xEnableWanted := TRUE; Warning.uiCode := UINT#1; Warning.udiSequence := Warning.udiSequence + UDINT#1;
			ELSE xEnabled := TRUE; END_IF;
			xCommandAccepted := TRUE;
		END_IF;
	UINT#2:
		IF Status.xDisableAllowed THEN
			xEnableWanted := FALSE; xManualRun := FALSE;
			IF Signals.xRobotInteraction THEN xDisablePending := TRUE;
			ELSE
				xEnabled := FALSE; xTransport := FALSE;
				IF Memory.xOccupied OR xReserved THEN Memory.xRecoveryRequired := TRUE; END_IF;
			END_IF;
			xCommandAccepted := TRUE;
		END_IF;
	UINT#3:
		IF Status.xConfirmAllowed THEN
			IF Memory.xOccupied AND (Memory.Part.udiId <> UDINT#0) THEN
				stRemoved := Memory.Part; stRemoved.uiState := UINT#8; F_GEOMETRY_EVENT(Call := stRemoved);
				IF (stRemoved.uiMachine >= UINT#1) AND (stRemoved.uiMachine <= UINT#3) THEN
					IF GVL_GEOMETRY_CONTROL.astCalls[stRemoved.uiMachine].udiId = stRemoved.udiId THEN
						GVL_GEOMETRY_CONTROL.astCalls[stRemoved.uiMachine] := stRemoved;
					END_IF;
				END_IF;
			END_IF;
			Memory.xOccupied := FALSE; Memory.xAtEndSeen := FALSE; Memory.xRecoveryRequired := FALSE;
			Memory.Part.udiId := UDINT#0; Memory.Part.uiMachine := UINT#0; Memory.Part.uiProductType := UINT#0;
			// Самостоятельное подтверждение состояния не включает станцию.
			xEnabled := xEnableWanted;
			xReserved := FALSE; xEnableWanted := FALSE; xCommandAccepted := TRUE;
			xSimulationEmptyConfirmed := xSimulation;
		END_IF;
	UINT#4:
		IF xEnableWanted OR Memory.xRecoveryRequired THEN
			xEnableWanted := FALSE; xEnabled := FALSE; xCommandAccepted := TRUE;
			Warning.uiCode := UINT#2; Warning.udiSequence := Warning.udiSequence + UDINT#1;
		END_IF;
	UINT#5:
		IF Status.xManualStartAllowed THEN
			xManualRun := TRUE; xCommandAccepted := TRUE;
			IF Memory.xOccupied THEN Memory.xRecoveryRequired := TRUE; xEnabled := FALSE; END_IF;
		END_IF;
	UINT#6:
		xManualRun := FALSE; xTransport := FALSE; xCommandAccepted := TRUE;
		IF Signals.xRobotInteraction THEN xDisablePending := TRUE;
		ELSIF Memory.xOccupied THEN Memory.xRecoveryRequired := TRUE; xEnabled := FALSE; END_IF;
	UINT#7:
		IF Status.xSimulationRemoveAllowed THEN
			xCommandAccepted := TRUE; xSimulationEmptyConfirmed := TRUE;
			xTransport := FALSE; xManualRun := FALSE;
		END_IF;
END_CASE;
IF (uiAction >= UINT#1) AND (uiAction <= UINT#7) AND NOT xCommandAccepted THEN xCommandRejected := TRUE; END_IF;
IF xDisablePending AND NOT Signals.xRobotInteraction THEN
	xEnabled := FALSE; xTransport := FALSE; xDisablePending := FALSE;
	IF Memory.xOccupied OR xReserved THEN Memory.xRecoveryRequired := TRUE; END_IF;
END_IF;

// Сброс привода — настоящий импульс. Внутренняя авария снимается после импульса,
// только при исчезновении входа. Занятость и требование восстановления сохраняются.
IF xReset AND NOT xResetSeen AND Status.xResetAllowed THEN xResetBusy := TRUE; END_IF;
xResetSeen := xReset;
tonReset(IN := xResetBusy, PT := tResetPulse);
xResetOutput := xResetBusy AND NOT tonReset.Q AND xSupported AND NOT xIoManual AND NOT xGlobalError;
IF xResetBusy AND tonReset.Q THEN
	xResetBusy := FALSE;
	IF NOT xDriveAlarm AND NOT xDriveRunning THEN Memory.dwAlarm := DWORD#0; Memory.xRobotStopLatched := FALSE; END_IF;
END_IF;

IF xTransport AND xPartAtEnd THEN
	Memory.xAtEndSeen := TRUE; xTransport := FALSE;
END_IF;
// В ручном режиме датчик никогда не останавливает привод.
xRunOutput := (xTransport OR xManualRun) AND NOT Signals.xRobotInteraction
	AND NOT xGlobalError AND xSupported AND NOT xIoManual AND NOT xDriveAlarm
	AND (Memory.dwAlarm = DWORD#0) AND NOT xResetBusy;
tonTransport(IN := xTransport AND xRunOutput, PT := tTransportScaled);
tonFeedback(IN := (xRunOutput <> xDriveRunning) AND NOT xResetBusy AND xSupported AND NOT xIoManual AND NOT xGlobalError, PT := tFeedbackScaled);
IF tonTransport.Q THEN Memory.dwAlarm := Memory.dwAlarm OR DWORD#2; END_IF;
IF tonFeedback.Q THEN Memory.dwAlarm := Memory.dwAlarm OR DWORD#4; END_IF;
IF Memory.dwAlarm <> DWORD#0 THEN
	xEnabled := FALSE; xEnableWanted := FALSE; xRunOutput := FALSE;
	xTransport := FALSE; xManualRun := FALSE; Memory.xRecoveryRequired := TRUE;
	IF Signals.xRobotInteraction THEN Memory.xRobotStopLatched := TRUE; END_IF;
END_IF;
tonRemoved(IN := Memory.xOccupied AND Memory.xAtEndSeen AND NOT xPartAtEnd
	AND xEnabled AND NOT Memory.xRecoveryRequired AND NOT xTransport AND NOT xManualRun
	AND NOT xDriveRunning AND NOT xReserved AND NOT Signals.xRobotInteraction
	AND (Memory.dwAlarm = DWORD#0) AND NOT xGlobalError, PT := T#3S);
// Явное изъятие в SIMULATION подтверждает пустоту всей ленты сразу.
// В NORMAL освобождение по датчику по-прежнему требует непрерывные 3 секунды.
IF tonRemoved.Q OR (xSimulationEmptyConfirmed AND Memory.xOccupied) THEN
	stRemoved := Memory.Part; stRemoved.uiState := UINT#8; F_GEOMETRY_EVENT(Call := stRemoved);
	IF (stRemoved.uiMachine >= UINT#1) AND (stRemoved.uiMachine <= UINT#3) THEN
		IF GVL_GEOMETRY_CONTROL.astCalls[stRemoved.uiMachine].udiId = stRemoved.udiId THEN
			GVL_GEOMETRY_CONTROL.astCalls[stRemoved.uiMachine] := stRemoved;
		END_IF;
	END_IF;
	Memory.xOccupied := FALSE; Memory.xAtEndSeen := FALSE;
	Memory.Part.udiId := UDINT#0; Memory.Part.uiMachine := UINT#0; Memory.Part.uiProductType := UINT#0;
END_IF;
IF xPartAtEnd AND NOT xSimulationEmptyConfirmed AND NOT Memory.xOccupied AND NOT xReserved THEN
	Memory.xRecoveryRequired := TRUE; xEnabled := FALSE;
END_IF;
IF xCommandRejected THEN Warning.uiCode := UINT#3; Warning.udiSequence := Warning.udiSequence + UDINT#1; END_IF;
Status.xEnabled := xEnabled;
Status.xReserved := xReserved;
// Виртуальный датчик снимается моделью на следующем скане после принятой команды.
Status.xPartAtEnd := xPartAtEnd AND NOT xSimulationEmptyConfirmed;
Status.xOccupied := Memory.xOccupied OR xReserved OR Memory.xRecoveryRequired OR Status.xPartAtEnd;
Status.xPartStored := Memory.xOccupied;
Status.xReady := xEnabled AND xConfigurationValid AND NOT Status.xOccupied AND NOT xDriveRunning
	AND (Memory.dwAlarm = DWORD#0) AND NOT xGlobalError AND xSupported AND NOT xIoManual AND NOT xResetBusy;
Status.xDriveRunning := xDriveRunning;
Status.xDriveAlarm := xDriveAlarm;
Status.xError := Memory.dwAlarm <> DWORD#0;
Status.xRobotStopRequired := Memory.xRobotStopLatched AND Status.xError;
Status.xResetBusy := xResetBusy;
Status.xConfirmationActive := xEnableWanted;
Status.xRecoveryRequired := Memory.xRecoveryRequired;
Status.xConfigured := xConfigurationValid;
Status.udiProducedPartsTotal := Memory.udiProducedPartsTotal;
Status.udiPartId := Memory.Part.udiId;
Status.uiMachine := Memory.Part.uiMachine;
Status.uiProductType := Memory.Part.uiProductType;
IF xSimulationEmptyConfirmed THEN Status.rTravel := REAL#0.0;
ELSIF xSimulation THEN Status.rTravel := rSimulationTravel;
ELSIF Memory.xAtEndSeen THEN Status.rTravel := REAL#1.0;
ELSIF xTransport THEN Status.rTravel := MIN(REAL#0.95, TIME_TO_REAL(tonTransport.ET) / TIME_TO_REAL(tTransportScaled));
ELSIF NOT Memory.xOccupied THEN Status.rTravel := REAL#0.0; END_IF;
IF Status.xError THEN Status.uiState := UINT#6;
ELSIF Memory.xRecoveryRequired THEN Status.uiState := UINT#5;
ELSIF xManualRun THEN Status.uiState := UINT#7;
ELSIF NOT xEnabled THEN Status.uiState := UINT#0;
ELSIF xReserved THEN Status.uiState := UINT#2;
ELSIF xTransport THEN Status.uiState := UINT#3;
ELSIF Memory.xOccupied THEN Status.uiState := UINT#4;
ELSE Status.uiState := UINT#1; END_IF;

END_FUNCTION_BLOCK

// Device/Application/FB/F_GEOMETRY_EVENT
FUNCTION F_GEOMETRY_EVENT : BOOL
VAR_INPUT
	Call : ST_GEOMETRY_CALL;
END_VAR
VAR
	uiIndex : UINT;
END_VAR

// Один PLC-скан, единый владелец номера. Поля записываются раньше Seq.
GVL_GEOMETRY_CONTROL.udiEventSequence := GVL_GEOMETRY_CONTROL.udiEventSequence + UDINT#1;
IF GVL_GEOMETRY_CONTROL.udiEventSequence = UDINT#0 THEN GVL_GEOMETRY_CONTROL.udiEventSequence := UDINT#1; END_IF;
uiIndex := UDINT_TO_UINT((GVL_GEOMETRY_CONTROL.udiEventSequence - UDINT#1) MOD UDINT#100) + UINT#1;
GVL_GEOMETRY_CONTROL.astEvents[uiIndex].udiSequence := UDINT#0;
GVL_GEOMETRY_CONTROL.astEvents[uiIndex].Call := Call;
GVL_GEOMETRY_CONTROL.astEvents[uiIndex].udiTimeMs := GVL_HMI.udiHmiCommandClockMs;
GVL_GEOMETRY_CONTROL.astEvents[uiIndex].uiEnvironment := GVL_GEOMETRY_CONTROL.uiEnvironment;
GVL_GEOMETRY_CONTROL.astEvents[uiIndex].udiSequence := GVL_GEOMETRY_CONTROL.udiEventSequence;
F_GEOMETRY_EVENT := TRUE;

END_FUNCTION

// Device/Application/FB/FB_GEOMETRY_CONTROL_SIMULATION
FUNCTION_BLOCK FB_GEOMETRY_CONTROL_SIMULATION
VAR_INPUT
	xInitialize : BOOL;
	xRun : BOOL;
	xReset : BOOL;
	xDeposited : BOOL;
	udiPartId : UDINT;
	xRemove : BOOL;
	xAlarm : BOOL;
	uiTimeFactor : UINT := UINT#1;
	tTravel : TIME := T#6S;
END_VAR
VAR_OUTPUT
	xDriveRunning : BOOL;
	xDriveAlarm : BOOL;
	xPartAtEnd : BOOL;
	rTravel : REAL;
END_VAR
VAR
	xPart : BOOL;
	udiSeenDeposit : UDINT;
	udiPreviousClock : UDINT;
	udiDeltaMs : UDINT;
	rElapsedMs : REAL;
END_VAR

IF xInitialize THEN
	xPart := FALSE; xPartAtEnd := FALSE; rTravel := REAL#0.0; udiSeenDeposit := UDINT#0;
	rElapsedMs := REAL#0.0; udiPreviousClock := GVL_HMI.udiHmiCommandClockMs;
END_IF;

// Накопленный путь сохраняется при останове и аварии. TON с IN=FALSE его теряет.
udiDeltaMs := MIN(UDINT#1000, GVL_HMI.udiHmiCommandClockMs - udiPreviousClock);
udiPreviousClock := GVL_HMI.udiHmiCommandClockMs;
IF xDeposited AND (udiPartId <> UDINT#0) AND (udiPartId <> udiSeenDeposit) THEN
	xPart := TRUE; xPartAtEnd := FALSE; rTravel := REAL#0.0; rElapsedMs := REAL#0.0; udiSeenDeposit := udiPartId;
END_IF;
IF xRemove THEN xPart := FALSE; xPartAtEnd := FALSE; rTravel := REAL#0.0; rElapsedMs := REAL#0.0; END_IF;
xDriveAlarm := xAlarm; // Сброс выхода не снимает удерживаемую физическую причину.
xDriveRunning := xRun AND NOT xDriveAlarm;
IF xPart AND NOT xPartAtEnd AND xDriveRunning THEN
	rElapsedMs := rElapsedMs + UDINT_TO_REAL(udiDeltaMs) * UINT_TO_REAL(MAX(UINT#1, uiTimeFactor));
	rTravel := MIN(REAL#1.0, rElapsedMs / MAX(REAL#1.0, TIME_TO_REAL(tTravel)));
	IF rTravel >= REAL#1.0 THEN xPartAtEnd := TRUE; END_IF;
END_IF;

END_FUNCTION_BLOCK

// Device/Application/FB/FB_DI_FILTER
FUNCTION_BLOCK FB_DI_FILTER
VAR_INPUT
	xEnable : BOOL;
	xInput : BOOL;
	tRise : TIME := T#20MS; // Стабильный 0 -> 1
	tFall : TIME := T#20MS; // Стабильный 1 -> 0
END_VAR
VAR_OUTPUT
	xFiltered : BOOL;
END_VAR
VAR
	tonRise : TON;
	tonFall : TON;
END_VAR

// Каждая смена направления сбрасывает противоположный таймер. Короткие
// выбросы не накапливаются. При нулевом времени уровень меняется в этом скане.
IF NOT xEnable THEN
	xFiltered := FALSE;
END_IF;
tonRise(IN := xEnable AND xInput AND NOT xFiltered, PT := tRise);
tonFall(IN := xEnable AND NOT xInput AND xFiltered, PT := tFall);
IF xEnable THEN
	IF xInput AND ((tRise = T#0MS) OR tonRise.Q) THEN
		xFiltered := TRUE;
	ELSIF NOT xInput AND ((tFall = T#0MS) OR tonFall.Q) THEN
		xFiltered := FALSE;
	END_IF;
END_IF;

END_FUNCTION_BLOCK

// Device/Application/FB/FB_AXIS
FUNCTION_BLOCK FB_Axis
VAR_INPUT
	FaultRequest : ST_AXIS_FAULT_REQUEST; // Единый контракт диагностической инъекции
	xResetPermit : BOOL; // Общий сброс разрешён ручным режимом и остановленной ячейкой
END_VAR
VAR_OUTPUT
	FaultStatus : ST_FAULT_INJECTION_STATUS; // Состояние инжектора для HMI
END_VAR
VAR_IN_OUT
    Axis     : AXIS_REF_SM3;   // ссылка на ось SoftMotion
    AxisData : ST_AXIS;        // все данные оси (команды, параметры, статусы)
END_VAR

VAR CONSTANT
    // ==================================================
    // Ошибки оси, MC-блоков и SoftMotion
    // ==================================================
    AXE_MC_POWER_ERROR       : DWORD := DWORD#16#00000001; // Ошибка MC_Power
    AXE_MC_RESET_ERROR       : DWORD := DWORD#16#00000002; // Ошибка MC_Reset
    AXE_MC_STOP_ERROR        : DWORD := DWORD#16#00000004; // Ошибка MC_Stop
    AXE_MC_JOG_ERROR         : DWORD := DWORD#16#00000008; // Ошибка MC_Jog
    AXE_MC_HOME_ERROR        : DWORD := DWORD#16#00000010; // Ошибка MC_Home
    AXE_MC_MOVE_ABS_ERROR    : DWORD := DWORD#16#00000020; // Ошибка абсолютного перемещения
    AXE_MC_MOVE_REL_ERROR    : DWORD := DWORD#16#00000040; // Ошибка относительного перемещения
    AXE_READ_POS_ERROR       : DWORD := DWORD#16#00000080; // Ошибка чтения позиции
    AXE_READ_STATUS_ERROR    : DWORD := DWORD#16#00000100; // Ошибка чтения статуса
    AXE_ERRORSTOP            : DWORD := DWORD#16#00000200; // Ось находится в ErrorStop
    AXE_FB_ERROR_OCCURRED    : DWORD := DWORD#16#00000400; // SoftMotion сообщил внутреннюю ошибку
    AXE_COMMAND_ABORTED      : DWORD := DWORD#16#00000800; // Команда движения прервана
    AXE_UNKNOWN_ACTUAL_ERROR : DWORD := DWORD#16#00001000; // Неизвестная текущая ошибка
    AXE_DRIVE_AXIS_ERROR     : DWORD := DWORD#16#00002000; // Ошибка привода
    AXE_POWER_FEEDBACK_LOST  : DWORD := DWORD#16#00004000; // Потеря силовой готовности при активной команде питания


    // ==================================================
    // Логические ошибки блока
    // ==================================================
    LOG_POWER_PERMIT_LOST    : DWORD := DWORD#16#00000001; // Снято разрешение питания
    LOG_GLOBAL_DURING_POWER  : DWORD := DWORD#16#00000002; // Глобальная ошибка при включении
    LOG_GLOBAL_DURING_READY  : DWORD := DWORD#16#00000004; // Глобальная ошибка в готовности
    LOG_GLOBAL_DURING_MOTION : DWORD := DWORD#16#00000008; // Глобальная ошибка при движении
    LOG_JOG_CONFLICT         : DWORD := DWORD#16#00000010; // Одновременно заданы Jog+ и Jog-
    LOG_MOVE_ABS_NOT_HOMED   : DWORD := DWORD#16#00000020; // Абсолютное движение без поиска дома
    LOG_MOVE_REL_NOT_HOMED   : DWORD := DWORD#16#00000040; // Относительное движение без поиска дома
    LOG_STEP_TIMEOUT         : DWORD := DWORD#16#00000080; // Превышено время шага
    LOG_UNKNOWN_STEP         : DWORD := DWORD#16#00000100; // Неизвестный шаг автомата

    // ==================================================
    // Предупреждения блока
    // ==================================================
    WRN_NO_POWER_PERMIT : DWORD := DWORD#16#00000001; // Нет разрешения подачи питания
    WRN_RESET_GLOBAL_ERROR   : UINT := 2; // Сброс не выполнен из-за глобальной ошибки
    WRN_RESET_MC_ERROR       : UINT := 3; // MC_Reset завершился ошибкой
    WRN_RESET_TIMEOUT        : UINT := 4; // Превышено время сброса
    WRN_RESET_AXIS_ACTIVE    : UINT := 5; // Физическая ошибка оси осталась активной
    WRN_RESET_AXIS_LATCHED   : UINT := 6; // Защёлкнутая ошибка оси не была очищена
    WRN_RESET_LOGICAL_ACTIVE : UINT := 7; // Логическая ошибка оси не была очищена
	WRN_SIM_ERROR_NOT_ALLOWED : UINT := 8; // Тестовый конфликт Jog запрещён состоянием оси

END_VAR

VAR
	lrEffectiveVelocity : LREAL;
	lrEffectiveAcceleration : LREAL;
	lrEffectiveDeceleration : LREAL;
	lrEffectiveJerk : LREAL;
    // Триггеры на команды
    rtEnable            : R_TRIG; // Фронт команды включения
    rtDisable           : R_TRIG; // Фронт команды отключения
    rtResetAllError     : R_TRIG; // Фронт общего сброса
    rtResetAxisError    : R_TRIG; // Фронт сброса привода
    rtResetLogicalError : R_TRIG; // Фронт сброса логики
    rtStop              : R_TRIG; // Фронт команды остановки
    rtHome              : R_TRIG; // Фронт команды поиска дома
    rtMoveAbsolute      : R_TRIG; // Фронт абсолютного перемещения
    rtMoveRelative      : R_TRIG; // Фронт относительного перемещения

    // Экземпляры MC-блоков
    fbPower        : MC_Power; // Управление питанием привода
    fbReset        : MC_Reset; // Сброс ошибки привода
    fbStop         : MC_Stop; // Контролируемая остановка
    fbJog          : MC_Jog; // Толчковое движение
    fbHome         : MC_Home; // Поиск домашней позиции
    fbMoveAbsolute : MC_MoveAbsolute; // Абсолютное перемещение
    fbMoveRelative : MC_MoveRelative; // Относительное перемещение
    fbReadPosition : MC_ReadActualPosition; // Чтение текущей позиции
    fbReadStatus   : MC_ReadStatus; // Чтение состояния оси
    fbReadAxisError: MC_ReadAxisError; // Чтение кода ошибки привода

    // Внутренние управляющие флаги 
    xPowerRequest    : BOOL; // Защёлкнутый запрос питания
    xResetExecute    : BOOL; // Выполняется сброс привода
    xStopExecute     : BOOL; // Выполняется остановка
    xHomeExecute     : BOOL; // Выполняется поиск дома
    xMoveAbsExecute  : BOOL; // Выполняется абсолютное перемещение
    xMoveRelExecute  : BOOL; // Выполняется относительное перемещение
    xJogForwardExec  : BOOL; // Выполняется Jog в положительную сторону
    xJogBackwardExec : BOOL; // Выполняется Jog в отрицательную сторону

    // Для таймера шага
    iPrevStep        : E_AXIS_STATE := E_AXIS_STATE.DISABLED; // Предыдущий шаг автомата
    xStepChanged     : BOOL; // Шаг изменился в текущем цикле
    xStepTimerEnable : BOOL; // Разрешение таймера шага
    tonStep          : TON; // Таймер времени на шаге
    tonStepTimeout   : TON; // Таймер превышения времени шага
    tonPowerFeedbackLoss : TON; // Контроль неожиданного снятия силовой готовности
    xPowerFeedbackExpected : BOOL; // Текущее состояние требует сохранения питания

    // Для удержания предупреждений
    tpWarningHold : TP; // Удержание предупреждения для отображения
    xWarningPulse : BOOL; // Импульс нового предупреждения

    // Вспомогательные флаги для сброса
    xDoResetAxis    : BOOL; // Требуется сброс ошибок привода
    xDoResetLogical : BOOL; // Требуется сброс логических ошибок
    xNeedMcReset    : BOOL; // Требуется вызов MC_Reset
    uiResetWarningCode : UINT; // Причина неуспешного сброса текущего цикла

    // Актуальная ошибка оси (на основе MC-блоков)
    xAxisErrorActual : BOOL; // Текущая ошибка по выходам MC-блоков
	fbFaultInjector : FB_AXIS_FAULT_INJECTOR; // Безопасный источник логической ошибки Jog
	xFaultAllowed   : BOOL; // Условия теста, рассчитанные владельцем оси
END_VAR

// Коэффициент симуляции не изменяет динамику осей робота.
// Скорость, ускорение, замедление и jerk задаются пользователем в настройках осей.
lrEffectiveVelocity := AxisData.MotionParam.lrVelocity;
lrEffectiveAcceleration := AxisData.MotionParam.lrAcceleration;
lrEffectiveDeceleration := AxisData.MotionParam.lrDeceleration;
lrEffectiveJerk := AxisData.MotionParam.lrJerk;

// ======================================================
// 1. ФРОНТЫ (триггеры на команды из структуры)
// ======================================================
rtEnable(CLK := AxisData.Command.xEnable);
rtDisable(CLK := AxisData.Command.xDisable);
rtResetAllError(CLK := AxisData.Command.xResetAllError);
rtResetAxisError(CLK := AxisData.Command.xResetAxisError);
rtResetLogicalError(CLK := AxisData.Command.xResetLogicalError);
rtStop(CLK := AxisData.Command.xStop);
rtHome(CLK := AxisData.Command.xHome);
rtMoveAbsolute(CLK := AxisData.Command.xMoveAbsolute);
rtMoveRelative(CLK := AxisData.Command.xMoveRelative);

// ======================================================
// 2. СТАТУСЫ ОТ MC-БЛОКОВ (запись в структуру)
// ======================================================
AxisData.Status.xPowerStageOn := fbPower.bRegulatorRealState;
AxisData.Status.xDriveStartOn := fbPower.bDriveStartRealState;
AxisData.Status.xPowered := fbPower.Status
	AND AxisData.Status.xPowerStageOn
	AND AxisData.Status.xDriveStartOn;
AxisData.Status.xPowerOff := NOT AxisData.Status.xPowerStageOn
	AND NOT AxisData.Status.xDriveStartOn;

AxisData.Status.xLocalError :=
    fbPower.Error OR
    fbReset.Error OR
    fbStop.Error OR
    fbJog.Error OR
    fbHome.Error OR
    fbMoveAbsolute.Error OR
    fbMoveRelative.Error OR
    fbReadPosition.Error OR
    fbReadStatus.Error OR
    fbReadStatus.Errorstop OR
    fbReadStatus.FBErrorOccured;

AxisData.Status.xMotionBusy :=
    fbStop.Busy OR
    fbJog.Busy OR
    fbHome.Busy OR
    fbMoveAbsolute.Busy OR
    fbMoveRelative.Busy;

// MC_Reset нужен только для аппаратных/SoftMotion ошибок
xNeedMcReset := fbReadStatus.Errorstop OR fbReadStatus.FBErrorOccured OR fbReadAxisError.AxisError;

AxisData.Error.dwAxisError := AxisData.Error.dwAxisErrorActual OR AxisData.Error.dwAxisErrorLatched;
AxisData.Error.dwLogicalError := AxisData.Error.dwLogicalErrorLatched;
AxisData.Error.dwAllError := AxisData.Error.dwAxisError OR AxisData.Error.dwLogicalError;

// ======================================================
// 3. ЗНАЧЕНИЯ ПО УМОЛЧАНИЮ ДЛЯ ИСПОЛНИТЕЛЬНЫХ ФЛАГОВ
// ======================================================
xResetExecute    := FALSE;
xStopExecute     := FALSE;
xHomeExecute     := FALSE;
xMoveAbsExecute  := FALSE;
xMoveRelExecute  := FALSE;
xJogForwardExec  := FALSE;
xJogBackwardExec := FALSE;

AxisData.Status.xDone := FALSE;
xWarningPulse := FALSE;
uiResetWarningCode := UINT#0;

// MC_Power не обязан выставлять Error при отказе интерфейса привода. Например,
// окончание demo-лицензии SoftMotion снимает реальные Regulator/DriveStart,
// но оставляет AxisError и FBError пустыми. Контролируем поэтому сам факт
// исчезновения силовой готовности при сохраняющемся запросе питания.
xPowerFeedbackExpected := xPowerRequest
	AND AxisData.Command.xPowerPermit
	AND ((AxisData.Diag.iStep = E_AXIS_STATE.READY)
		OR (AxisData.Diag.iStep = E_AXIS_STATE.JOGGING)
		OR (AxisData.Diag.iStep = E_AXIS_STATE.JOG_DECELERATING)
		OR (AxisData.Diag.iStep = E_AXIS_STATE.HOMING)
		OR (AxisData.Diag.iStep = E_AXIS_STATE.MOVE_ABSOLUTE)
		OR (AxisData.Diag.iStep = E_AXIS_STATE.MOVE_RELATIVE)
		OR (AxisData.Diag.iStep = E_AXIS_STATE.STOPPING)
		OR (AxisData.Diag.iStep = E_AXIS_STATE.STOP_RELEASE));
tonPowerFeedbackLoss(
	IN := xPowerFeedbackExpected AND NOT AxisData.Status.xPowered,
	PT := AxisData.Timeouts.tPowerFeedbackLossTimeout
);
IF tonPowerFeedbackLoss.Q
AND (AxisData.Diag.iStep <> E_AXIS_STATE.ERROR_RESET_MANAGER) THEN
	AxisData.Error.dwAxisErrorLatched :=
		AxisData.Error.dwAxisErrorLatched OR AXE_POWER_FEEDBACK_LOST;
	AxisData.Diag.iLastErrorStep := TO_INT(AxisData.Diag.iStep);
	AxisData.Diag.iStep := E_AXIS_STATE.ERROR_RESET_MANAGER;
END_IF;

// Конфликт Jog проверяется автоматом до вызова MC_Jog, поэтому тест не создаёт движения.
xFaultAllowed := (AxisData.Diag.iStep = E_AXIS_STATE.READY)
	AND NOT AxisData.Command.xGlobalError
	AND NOT AxisData.Status.xError
	AND NOT AxisData.Status.xMotionBusy
	AND NOT AxisData.Command.xJogPositive
	AND NOT AxisData.Command.xJogNegative
	AND NOT AxisData.Command.xHome
	AND NOT AxisData.Command.xMoveAbsolute
	AND NOT AxisData.Command.xMoveRelative;

fbFaultInjector(
	Request := FaultRequest,
	xOwnerAllowed := xFaultAllowed
);
FaultStatus := fbFaultInjector.Status;

IF fbFaultInjector.Status.xRejected THEN
	AxisData.Diag.sWarningText := 'Simulated Jog conflict is not allowed';
	AxisData.Diag.stWarning.uiCode := WRN_SIM_ERROR_NOT_ALLOWED;
	AxisData.Diag.stWarning.udiSequence := AxisData.Diag.stWarning.udiSequence + UDINT#1;
	IF AxisData.Diag.stWarning.udiSequence = UDINT#0 THEN
		AxisData.Diag.stWarning.udiSequence := UDINT#1;
	END_IF;
	xWarningPulse := TRUE;
END_IF;

// ======================================================
// 4. КОНЕЧНЫЙ АВТОМАТ (используем перечисление E_AXIS_STATE)
// ======================================================
CASE AxisData.Diag.iStep OF

    // --------------------------------------------------
    E_AXIS_STATE.DISABLED:
    // --------------------------------------------------
        AxisData.Diag.sStepName := 'DISABLED';
        AxisData.Diag.sWaitReason := 'Waiting Enable command';
        AxisData.Diag.tStepPreset := T#0S;

        xPowerRequest := FALSE;
        AxisData.Status.xHomed := FALSE;

        IF AxisData.Status.xError THEN
            AxisData.Diag.iStep := E_AXIS_STATE.ERROR_RESET_MANAGER;

        ELSIF rtEnable.Q AND NOT AxisData.Command.xPowerPermit THEN
            AxisData.Error.dwWarningLatched :=
                AxisData.Error.dwWarningLatched OR WRN_NO_POWER_PERMIT;
            AxisData.Diag.sWarningText := 'Power permit is not active';
            AxisData.Diag.stWarning.uiCode := UINT#1;
            AxisData.Diag.stWarning.udiSequence := AxisData.Diag.stWarning.udiSequence + UDINT#1;
            IF AxisData.Diag.stWarning.udiSequence = UDINT#0 THEN
                AxisData.Diag.stWarning.udiSequence := UDINT#1;
            END_IF;
            xWarningPulse := TRUE;
            AxisData.Diag.sWaitReason := 'Power permit missing';

        ELSIF NOT AxisData.Command.xPowerPermit THEN
            AxisData.Diag.sWaitReason := 'Power permit missing';

        ELSIF rtEnable.Q THEN
            xPowerRequest := TRUE;
            AxisData.Diag.iStep := E_AXIS_STATE.POWERING;
        END_IF;

    // --------------------------------------------------
    E_AXIS_STATE.POWERING:
    // --------------------------------------------------
        AxisData.Diag.sStepName := 'POWERING';
        AxisData.Diag.sWaitReason := 'Waiting MC_Power.Status';
        AxisData.Diag.tStepPreset := AxisData.Timeouts.tPowerTimeout;

        xPowerRequest := TRUE;

        IF NOT AxisData.Command.xPowerPermit THEN
            xPowerRequest := FALSE;
            AxisData.Error.dwLogicalErrorLatched :=
                AxisData.Error.dwLogicalErrorLatched OR LOG_POWER_PERMIT_LOST;
            AxisData.Diag.iLastErrorStep := TO_INT(AxisData.Diag.iStep);
            AxisData.Diag.iStep := E_AXIS_STATE.ERROR_RESET_MANAGER;

        ELSIF AxisData.Command.xGlobalError THEN
            xPowerRequest := FALSE;
            AxisData.Error.dwLogicalErrorLatched :=
                AxisData.Error.dwLogicalErrorLatched OR LOG_GLOBAL_DURING_POWER;
            AxisData.Diag.iLastErrorStep := TO_INT(AxisData.Diag.iStep);
            AxisData.Diag.iStep := E_AXIS_STATE.ERROR_RESET_MANAGER;

        ELSIF fbPower.Error THEN
            xPowerRequest := FALSE;
            AxisData.Error.dwAxisErrorLatched :=
                AxisData.Error.dwAxisErrorLatched OR AXE_MC_POWER_ERROR;
            AxisData.Diag.udiLastErrorID := TO_UDINT(fbPower.ErrorID);
            AxisData.Diag.iLastErrorStep := TO_INT(AxisData.Diag.iStep);
            AxisData.Diag.iStep := E_AXIS_STATE.ERROR_RESET_MANAGER;

        // READY допустим только после подтверждения всех трёх признаков:
        // MC_Power.Status, силовая ступень и снятый quickstop.
        ELSIF AxisData.Status.xPowered THEN
            AxisData.Diag.iStep := E_AXIS_STATE.READY;

        ELSIF rtDisable.Q THEN
            xPowerRequest := FALSE;
            AxisData.Diag.iStep := E_AXIS_STATE.POWERING_DOWN;
        END_IF;

    // --------------------------------------------------
    E_AXIS_STATE.POWERING_DOWN:
    // --------------------------------------------------
        AxisData.Diag.sStepName := 'POWERING_DOWN';
        AxisData.Diag.sWaitReason := 'Waiting drive power feedback off';
        AxisData.Diag.tStepPreset := AxisData.Timeouts.tPowerTimeout;

        xPowerRequest := FALSE;

        IF fbPower.Error THEN
            AxisData.Error.dwAxisErrorLatched :=
                AxisData.Error.dwAxisErrorLatched OR AXE_MC_POWER_ERROR;
            AxisData.Diag.udiLastErrorID := TO_UDINT(fbPower.ErrorID);
            AxisData.Diag.iLastErrorStep := TO_INT(AxisData.Diag.iStep);
            AxisData.Diag.iStep := E_AXIS_STATE.ERROR_RESET_MANAGER;

        ELSIF AxisData.Status.xPowerOff THEN
            AxisData.Diag.iStep := E_AXIS_STATE.DISABLED;
        END_IF;

    // --------------------------------------------------
    E_AXIS_STATE.READY:
    // --------------------------------------------------
        AxisData.Diag.sStepName := 'READY';
        AxisData.Diag.sWaitReason := 'Waiting command';
        AxisData.Diag.tStepPreset := T#0S;

        xPowerRequest := TRUE;

        IF NOT AxisData.Command.xPowerPermit THEN
            xPowerRequest := FALSE;
            AxisData.Diag.iStep := E_AXIS_STATE.POWERING_DOWN;

        ELSIF rtDisable.Q THEN
            xPowerRequest := FALSE;
            AxisData.Diag.iStep := E_AXIS_STATE.POWERING_DOWN;

        ELSIF AxisData.Command.xGlobalError THEN
            AxisData.Error.dwLogicalErrorLatched :=
                AxisData.Error.dwLogicalErrorLatched OR LOG_GLOBAL_DURING_READY;
            AxisData.Diag.iLastErrorStep := TO_INT(AxisData.Diag.iStep);
            AxisData.Diag.iStep := E_AXIS_STATE.ERROR_RESET_MANAGER;

        ELSIF xAxisErrorActual THEN
            AxisData.Error.dwAxisErrorLatched :=
                AxisData.Error.dwAxisErrorLatched OR AxisData.Error.dwAxisErrorActual;
            AxisData.Diag.iLastErrorStep := TO_INT(AxisData.Diag.iStep);
            AxisData.Diag.iStep := E_AXIS_STATE.ERROR_RESET_MANAGER;

        ELSIF fbFaultInjector.xJogConflict
		OR (AxisData.Command.xJogPositive AND AxisData.Command.xJogNegative) THEN
            AxisData.Error.dwLogicalErrorLatched :=
                AxisData.Error.dwLogicalErrorLatched OR LOG_JOG_CONFLICT;
            AxisData.Diag.iLastErrorStep := TO_INT(AxisData.Diag.iStep);
            AxisData.Diag.iStep := E_AXIS_STATE.ERROR_RESET_MANAGER;

        ELSIF AxisData.Command.xJogPositive OR AxisData.Command.xJogNegative THEN
            AxisData.Diag.iStep := E_AXIS_STATE.JOGGING;

        ELSIF rtHome.Q THEN
            AxisData.Diag.iStep := E_AXIS_STATE.HOMING;

        ELSIF rtMoveAbsolute.Q THEN
            IF AxisData.Status.xHomed THEN
                AxisData.Diag.iStep := E_AXIS_STATE.MOVE_ABSOLUTE;
            ELSE
                AxisData.Error.dwLogicalErrorLatched :=
                    AxisData.Error.dwLogicalErrorLatched OR LOG_MOVE_ABS_NOT_HOMED;
                AxisData.Diag.iLastErrorStep := TO_INT(AxisData.Diag.iStep);
                AxisData.Diag.iStep := E_AXIS_STATE.ERROR_RESET_MANAGER;
            END_IF;

        ELSIF rtMoveRelative.Q THEN
            IF AxisData.Status.xHomed THEN
                AxisData.Diag.iStep := E_AXIS_STATE.MOVE_RELATIVE;
            ELSE
                AxisData.Error.dwLogicalErrorLatched :=
                    AxisData.Error.dwLogicalErrorLatched OR LOG_MOVE_REL_NOT_HOMED;
                AxisData.Diag.iLastErrorStep := TO_INT(AxisData.Diag.iStep);
                AxisData.Diag.iStep := E_AXIS_STATE.ERROR_RESET_MANAGER;
            END_IF;
        END_IF;

    // --------------------------------------------------
    E_AXIS_STATE.JOGGING:
    // --------------------------------------------------
        AxisData.Diag.sStepName := 'JOGGING';
        AxisData.Diag.sWaitReason := 'Jog active';
        AxisData.Diag.tStepPreset := T#0S;

        xPowerRequest := TRUE;
        xJogForwardExec  := AxisData.Command.xJogPositive AND NOT AxisData.Command.xJogNegative;
        xJogBackwardExec := AxisData.Command.xJogNegative AND NOT AxisData.Command.xJogPositive;

        IF NOT AxisData.Command.xPowerPermit THEN
            xJogForwardExec := FALSE;
            xJogBackwardExec := FALSE;
            AxisData.Error.dwLogicalErrorLatched :=
                AxisData.Error.dwLogicalErrorLatched OR LOG_POWER_PERMIT_LOST;
            AxisData.Diag.iLastErrorStep := TO_INT(AxisData.Diag.iStep);
            AxisData.Diag.iStep := E_AXIS_STATE.STOPPING;

        ELSIF AxisData.Command.xGlobalError THEN
            xJogForwardExec := FALSE;
            xJogBackwardExec := FALSE;
            AxisData.Error.dwLogicalErrorLatched :=
                AxisData.Error.dwLogicalErrorLatched OR LOG_GLOBAL_DURING_MOTION;
            AxisData.Diag.iLastErrorStep := TO_INT(AxisData.Diag.iStep);
            AxisData.Diag.iStep := E_AXIS_STATE.STOPPING;

        ELSIF xAxisErrorActual THEN
            xJogForwardExec := FALSE;
            xJogBackwardExec := FALSE;
            AxisData.Error.dwAxisErrorLatched :=
                AxisData.Error.dwAxisErrorLatched OR AxisData.Error.dwAxisErrorActual;
            AxisData.Diag.iLastErrorStep := TO_INT(AxisData.Diag.iStep);
            // SoftMotion уже перевёл ось в ErrorStop и выполнил error ramp.
            // MC_Stop в этом состоянии создаёт вторичную ошибку "axis is in errorstop".
            AxisData.Diag.iStep := E_AXIS_STATE.ERROR_RESET_MANAGER;

        ELSIF rtStop.Q THEN
            xJogForwardExec := FALSE;
            xJogBackwardExec := FALSE;
            AxisData.Diag.iStep := E_AXIS_STATE.STOPPING;

        ELSIF AxisData.Command.xJogPositive AND AxisData.Command.xJogNegative THEN
            xJogForwardExec := FALSE;
            xJogBackwardExec := FALSE;
            AxisData.Error.dwLogicalErrorLatched :=
                AxisData.Error.dwLogicalErrorLatched OR LOG_JOG_CONFLICT;
            AxisData.Diag.iLastErrorStep := TO_INT(AxisData.Diag.iStep);
            AxisData.Diag.iStep := E_AXIS_STATE.STOPPING;

        ELSIF NOT AxisData.Command.xJogPositive AND NOT AxisData.Command.xJogNegative THEN
            xJogForwardExec := FALSE;
            xJogBackwardExec := FALSE;
            AxisData.Diag.iStep := E_AXIS_STATE.JOG_DECELERATING;
        END_IF;

    // --------------------------------------------------
    E_AXIS_STATE.JOG_DECELERATING:
    // --------------------------------------------------
        AxisData.Diag.sStepName := 'JOG_DECELERATING';
        AxisData.Diag.sWaitReason := 'Waiting MC_Jog controlled deceleration';
        AxisData.Diag.tStepPreset := T#0S;

        xPowerRequest := TRUE;
        xJogForwardExec := FALSE;
        xJogBackwardExec := FALSE;

        IF NOT AxisData.Command.xPowerPermit THEN
            AxisData.Error.dwLogicalErrorLatched :=
                AxisData.Error.dwLogicalErrorLatched OR LOG_POWER_PERMIT_LOST;
            AxisData.Diag.iLastErrorStep := TO_INT(AxisData.Diag.iStep);
            AxisData.Diag.iStep := E_AXIS_STATE.STOPPING;

        ELSIF AxisData.Command.xGlobalError THEN
            AxisData.Error.dwLogicalErrorLatched :=
                AxisData.Error.dwLogicalErrorLatched OR LOG_GLOBAL_DURING_MOTION;
            AxisData.Diag.iLastErrorStep := TO_INT(AxisData.Diag.iStep);
            AxisData.Diag.iStep := E_AXIS_STATE.STOPPING;

        ELSIF xAxisErrorActual THEN
            AxisData.Error.dwAxisErrorLatched :=
                AxisData.Error.dwAxisErrorLatched OR AxisData.Error.dwAxisErrorActual;
            AxisData.Diag.iLastErrorStep := TO_INT(AxisData.Diag.iStep);
            AxisData.Diag.iStep := E_AXIS_STATE.ERROR_RESET_MANAGER;

        ELSIF rtStop.Q THEN
            AxisData.Diag.iStep := E_AXIS_STATE.STOPPING;

        ELSIF AxisData.Command.xJogPositive AND AxisData.Command.xJogNegative THEN
            AxisData.Error.dwLogicalErrorLatched :=
                AxisData.Error.dwLogicalErrorLatched OR LOG_JOG_CONFLICT;
            AxisData.Diag.iLastErrorStep := TO_INT(AxisData.Diag.iStep);
            AxisData.Diag.iStep := E_AXIS_STATE.STOPPING;

        ELSIF AxisData.Command.xJogPositive OR AxisData.Command.xJogNegative THEN
            AxisData.Diag.iStep := E_AXIS_STATE.JOGGING;

        ELSIF NOT fbJog.Busy THEN
            AxisData.Status.xDone := TRUE;
            AxisData.Diag.iStep := E_AXIS_STATE.READY;
        END_IF;

    // --------------------------------------------------
    E_AXIS_STATE.HOMING:
    // --------------------------------------------------
        AxisData.Diag.sStepName := 'HOMING';
        AxisData.Diag.sWaitReason := 'Waiting MC_Home.Done';
        AxisData.Diag.tStepPreset := AxisData.Timeouts.tHomeTimeout;

        xPowerRequest := TRUE;
        xHomeExecute := TRUE;

        IF NOT AxisData.Command.xPowerPermit THEN
            xHomeExecute := FALSE;
            AxisData.Error.dwLogicalErrorLatched :=
                AxisData.Error.dwLogicalErrorLatched OR LOG_POWER_PERMIT_LOST;
            AxisData.Diag.iLastErrorStep := TO_INT(AxisData.Diag.iStep);
            AxisData.Diag.iStep := E_AXIS_STATE.STOPPING;

        ELSIF AxisData.Command.xGlobalError THEN
            xHomeExecute := FALSE;
            AxisData.Error.dwLogicalErrorLatched :=
                AxisData.Error.dwLogicalErrorLatched OR LOG_GLOBAL_DURING_MOTION;
            AxisData.Diag.iLastErrorStep := TO_INT(AxisData.Diag.iStep);
            AxisData.Diag.iStep := E_AXIS_STATE.STOPPING;

        ELSIF rtStop.Q THEN
            xHomeExecute := FALSE;
            AxisData.Diag.iStep := E_AXIS_STATE.STOPPING;

        ELSIF fbHome.Error THEN
            xHomeExecute := FALSE;
            AxisData.Error.dwAxisErrorLatched :=
                AxisData.Error.dwAxisErrorLatched OR AXE_MC_HOME_ERROR;
            AxisData.Diag.udiLastErrorID := TO_UDINT(fbHome.ErrorID);
            AxisData.Diag.iLastErrorStep := TO_INT(AxisData.Diag.iStep);
            AxisData.Diag.iStep := E_AXIS_STATE.ERROR_RESET_MANAGER;

        ELSIF fbHome.CommandAborted THEN
            xHomeExecute := FALSE;
            AxisData.Error.dwAxisErrorLatched :=
                AxisData.Error.dwAxisErrorLatched OR AXE_COMMAND_ABORTED;
            AxisData.Diag.udiLastErrorID := 3003;
            AxisData.Diag.iLastErrorStep := TO_INT(AxisData.Diag.iStep);
            AxisData.Diag.iStep := E_AXIS_STATE.ERROR_RESET_MANAGER;

        ELSIF xAxisErrorActual THEN
            xHomeExecute := FALSE;
            AxisData.Error.dwAxisErrorLatched :=
                AxisData.Error.dwAxisErrorLatched OR AxisData.Error.dwAxisErrorActual;
            AxisData.Diag.iLastErrorStep := TO_INT(AxisData.Diag.iStep);
            AxisData.Diag.iStep := E_AXIS_STATE.ERROR_RESET_MANAGER;

        ELSIF fbHome.Done THEN
            xHomeExecute := FALSE;
            AxisData.Status.xHomed := TRUE;
            AxisData.Status.xDone := TRUE;
            AxisData.Diag.iStep := E_AXIS_STATE.READY;
        END_IF;

    // --------------------------------------------------
    E_AXIS_STATE.MOVE_ABSOLUTE:
    // --------------------------------------------------
        AxisData.Diag.sStepName := 'MOVING_ABSOLUTE';
        AxisData.Diag.sWaitReason := 'Waiting MC_MoveAbsolute.Done';
        AxisData.Diag.tStepPreset := AxisData.Timeouts.tMoveTimeout;

        xPowerRequest := TRUE;
        xMoveAbsExecute := TRUE;

        IF NOT AxisData.Command.xPowerPermit THEN
            xMoveAbsExecute := FALSE;
            AxisData.Error.dwLogicalErrorLatched :=
                AxisData.Error.dwLogicalErrorLatched OR LOG_POWER_PERMIT_LOST;
            AxisData.Diag.iLastErrorStep := TO_INT(AxisData.Diag.iStep);
            AxisData.Diag.iStep := E_AXIS_STATE.STOPPING;

        ELSIF AxisData.Command.xGlobalError THEN
            xMoveAbsExecute := FALSE;
            AxisData.Error.dwLogicalErrorLatched :=
                AxisData.Error.dwLogicalErrorLatched OR LOG_GLOBAL_DURING_MOTION;
            AxisData.Diag.iLastErrorStep := TO_INT(AxisData.Diag.iStep);
            AxisData.Diag.iStep := E_AXIS_STATE.STOPPING;

        ELSIF rtStop.Q THEN
            xMoveAbsExecute := FALSE;
            AxisData.Diag.iStep := E_AXIS_STATE.STOPPING;

        ELSIF fbMoveAbsolute.Error THEN
            xMoveAbsExecute := FALSE;
            AxisData.Error.dwAxisErrorLatched :=
                AxisData.Error.dwAxisErrorLatched OR AXE_MC_MOVE_ABS_ERROR;
            AxisData.Diag.udiLastErrorID := TO_UDINT(fbMoveAbsolute.ErrorID);
            AxisData.Diag.iLastErrorStep := TO_INT(AxisData.Diag.iStep);
            AxisData.Diag.iStep := E_AXIS_STATE.ERROR_RESET_MANAGER;

        ELSIF fbMoveAbsolute.CommandAborted THEN
            xMoveAbsExecute := FALSE;
            AxisData.Error.dwAxisErrorLatched :=
                AxisData.Error.dwAxisErrorLatched OR AXE_COMMAND_ABORTED;
            AxisData.Diag.udiLastErrorID := 3003;
            AxisData.Diag.iLastErrorStep := TO_INT(AxisData.Diag.iStep);
            AxisData.Diag.iStep := E_AXIS_STATE.ERROR_RESET_MANAGER;

        ELSIF xAxisErrorActual THEN
            xMoveAbsExecute := FALSE;
            AxisData.Error.dwAxisErrorLatched :=
                AxisData.Error.dwAxisErrorLatched OR AxisData.Error.dwAxisErrorActual;
            AxisData.Diag.iLastErrorStep := TO_INT(AxisData.Diag.iStep);
            AxisData.Diag.iStep := E_AXIS_STATE.ERROR_RESET_MANAGER;

        ELSIF fbMoveAbsolute.Done THEN
            xMoveAbsExecute := FALSE;
            AxisData.Status.xDone := TRUE;
            AxisData.Diag.iStep := E_AXIS_STATE.READY;
        END_IF;

    // --------------------------------------------------
    E_AXIS_STATE.MOVE_RELATIVE:
    // --------------------------------------------------
        AxisData.Diag.sStepName := 'MOVING_RELATIVE';
        AxisData.Diag.sWaitReason := 'Waiting MC_MoveRelative.Done';
        AxisData.Diag.tStepPreset := AxisData.Timeouts.tMoveTimeout;

        xPowerRequest := TRUE;
        xMoveRelExecute := TRUE;

        IF NOT AxisData.Command.xPowerPermit THEN
            xMoveRelExecute := FALSE;
            AxisData.Error.dwLogicalErrorLatched :=
                AxisData.Error.dwLogicalErrorLatched OR LOG_POWER_PERMIT_LOST;
            AxisData.Diag.iLastErrorStep := TO_INT(AxisData.Diag.iStep);
            AxisData.Diag.iStep := E_AXIS_STATE.STOPPING;

        ELSIF AxisData.Command.xGlobalError THEN
            xMoveRelExecute := FALSE;
            AxisData.Error.dwLogicalErrorLatched :=
                AxisData.Error.dwLogicalErrorLatched OR LOG_GLOBAL_DURING_MOTION;
            AxisData.Diag.iLastErrorStep := TO_INT(AxisData.Diag.iStep);
            AxisData.Diag.iStep := E_AXIS_STATE.STOPPING;

        ELSIF rtStop.Q THEN
            xMoveRelExecute := FALSE;
            AxisData.Diag.iStep := E_AXIS_STATE.STOPPING;

        ELSIF fbMoveRelative.Error THEN
            xMoveRelExecute := FALSE;
            AxisData.Error.dwAxisErrorLatched :=
                AxisData.Error.dwAxisErrorLatched OR AXE_MC_MOVE_REL_ERROR;
            AxisData.Diag.udiLastErrorID := TO_UDINT(fbMoveRelative.ErrorID);
            AxisData.Diag.iLastErrorStep := TO_INT(AxisData.Diag.iStep);
            AxisData.Diag.iStep := E_AXIS_STATE.ERROR_RESET_MANAGER;

        ELSIF fbMoveRelative.CommandAborted THEN
            xMoveRelExecute := FALSE;
            AxisData.Error.dwAxisErrorLatched :=
                AxisData.Error.dwAxisErrorLatched OR AXE_COMMAND_ABORTED;
            AxisData.Diag.udiLastErrorID := 3003;
            AxisData.Diag.iLastErrorStep := TO_INT(AxisData.Diag.iStep);
            AxisData.Diag.iStep := E_AXIS_STATE.ERROR_RESET_MANAGER;

        ELSIF xAxisErrorActual THEN
            xMoveRelExecute := FALSE;
            AxisData.Error.dwAxisErrorLatched :=
                AxisData.Error.dwAxisErrorLatched OR AxisData.Error.dwAxisErrorActual;
            AxisData.Diag.iLastErrorStep := TO_INT(AxisData.Diag.iStep);
            AxisData.Diag.iStep := E_AXIS_STATE.ERROR_RESET_MANAGER;

        ELSIF fbMoveRelative.Done THEN 
            xMoveRelExecute := FALSE;
            AxisData.Status.xDone := TRUE;
            AxisData.Diag.iStep := E_AXIS_STATE.READY;
        END_IF;

    // --------------------------------------------------
    E_AXIS_STATE.STOPPING:
    // --------------------------------------------------
        AxisData.Diag.sStepName := 'STOPPING';
        AxisData.Diag.sWaitReason := 'Waiting MC_Stop.Done';
        AxisData.Diag.tStepPreset := AxisData.Timeouts.tStopTimeout;

        xPowerRequest := TRUE;
        xStopExecute := TRUE;

        IF fbStop.Error THEN
            xStopExecute := FALSE;
            AxisData.Error.dwAxisErrorLatched :=
                AxisData.Error.dwAxisErrorLatched OR AXE_MC_STOP_ERROR;
            AxisData.Diag.udiLastErrorID := TO_UDINT(fbStop.ErrorID);
            AxisData.Diag.iLastErrorStep := TO_INT(AxisData.Diag.iStep);
            AxisData.Diag.iStep := E_AXIS_STATE.ERROR_RESET_MANAGER;

        ELSIF fbStop.Done THEN
            AxisData.Status.xDone := TRUE;
            AxisData.Diag.iStep := E_AXIS_STATE.STOP_RELEASE;
        END_IF;

    // --------------------------------------------------
    E_AXIS_STATE.STOP_RELEASE:
    // --------------------------------------------------
        AxisData.Diag.sStepName := 'STOP_RELEASE';
        AxisData.Diag.sWaitReason := 'Releasing MC_Stop.Execute';
        AxisData.Diag.tStepPreset := T#1S;

        xPowerRequest := TRUE;
        xStopExecute := FALSE;

        IF NOT fbStop.Busy THEN
            IF AxisData.Command.xGlobalError OR
               (AxisData.Error.dwAxisErrorLatched <> DWORD#0) OR
               (AxisData.Error.dwLogicalErrorLatched <> DWORD#0) OR
               xAxisErrorActual
            THEN
                AxisData.Diag.iStep := E_AXIS_STATE.ERROR_RESET_MANAGER;
            ELSE
                AxisData.Diag.iStep := E_AXIS_STATE.READY;
            END_IF;
        END_IF;

    // --------------------------------------------------
    E_AXIS_STATE.ERROR_RESET_MANAGER:
    // --------------------------------------------------
        AxisData.Diag.sStepName := 'ERROR';
        AxisData.Diag.tStepPreset := T#0S;

        xResetExecute    := FALSE;
        xStopExecute     := FALSE;
        xHomeExecute     := FALSE;
        xMoveAbsExecute  := FALSE;
        xMoveRelExecute  := FALSE;
        xJogForwardExec  := FALSE;
        xJogBackwardExec := FALSE;

        IF AxisData.Timeouts.xDisableOnError THEN
            xPowerRequest := FALSE;
        ELSE
            xPowerRequest := AxisData.Command.xPowerPermit AND NOT xAxisErrorActual;
        END_IF;

        IF (AxisData.Error.dwAxisError = DWORD#0) AND
           (AxisData.Error.dwLogicalError = DWORD#0) AND
           NOT AxisData.Command.xGlobalError
        THEN
            AxisData.Diag.iStep := E_AXIS_STATE.DISABLED;

        ELSE
            IF AxisData.Command.xGlobalError THEN
                AxisData.Diag.sWaitReason := 'Waiting global error release';
            ELSIF (AxisData.Error.dwAxisError <> DWORD#0) AND
                  (AxisData.Error.dwLogicalError <> DWORD#0) THEN
                AxisData.Diag.sWaitReason := 'Waiting ResetAllError';
            ELSIF AxisData.Error.dwAxisError <> DWORD#0 THEN
                AxisData.Diag.sWaitReason := 'Waiting ResetAxisError or ResetAllError';
            ELSIF AxisData.Error.dwLogicalError <> DWORD#0 THEN
                AxisData.Diag.sWaitReason := 'Waiting ResetLogicalError or ResetAllError';
            ELSE
                AxisData.Diag.sWaitReason := 'Waiting reset';
            END_IF;

            IF rtResetAllError.Q AND xResetPermit THEN
                xDoResetAxis := TRUE;
                xDoResetLogical := TRUE;
                IF xNeedMcReset THEN
                    AxisData.Diag.iStep := E_AXIS_STATE.RESET_AXIS_ERROR;
                ELSE
                    AxisData.Diag.iStep := E_AXIS_STATE.RESET_FINISH;
                END_IF;

            ELSIF rtResetAxisError.Q THEN
                xDoResetAxis := TRUE;
                xDoResetLogical := FALSE;
                IF xNeedMcReset THEN
                    AxisData.Diag.iStep := E_AXIS_STATE.RESET_AXIS_ERROR;
                ELSE
                    AxisData.Diag.iStep := E_AXIS_STATE.RESET_FINISH;
                END_IF;

            ELSIF rtResetLogicalError.Q THEN
                xDoResetAxis := FALSE;
                xDoResetLogical := TRUE;
                AxisData.Diag.iStep := E_AXIS_STATE.RESET_FINISH;
            END_IF;
        END_IF;

    // --------------------------------------------------
    E_AXIS_STATE.RESET_AXIS_ERROR:
    // --------------------------------------------------
        AxisData.Diag.sStepName := 'RESET_AXIS_ERROR';
        AxisData.Diag.sWaitReason := 'Waiting MC_Reset.Done';
        AxisData.Diag.tStepPreset := AxisData.Timeouts.tResetTimeout;

        xPowerRequest := FALSE;
        xResetExecute := TRUE;

        IF fbReset.Error THEN
            AxisData.Diag.sWarningText := 'MC_Reset finished with error';
            uiResetWarningCode := WRN_RESET_MC_ERROR;
            xResetExecute := FALSE;
            AxisData.Error.dwAxisErrorLatched :=
                AxisData.Error.dwAxisErrorLatched OR AXE_MC_RESET_ERROR;
            AxisData.Diag.udiLastErrorID := TO_UDINT(fbReset.ErrorID);
            AxisData.Diag.iLastErrorStep := TO_INT(AxisData.Diag.iStep);
            AxisData.Diag.iStep := E_AXIS_STATE.ERROR_RESET_MANAGER;

        ELSIF fbReset.Done THEN
            xResetExecute := FALSE;
            AxisData.Diag.iStep := E_AXIS_STATE.RESET_RELEASE;
        END_IF;

    // --------------------------------------------------
    E_AXIS_STATE.RESET_RELEASE:
    // --------------------------------------------------
        AxisData.Diag.sStepName := 'RESET_RELEASE';
        AxisData.Diag.sWaitReason := 'Releasing MC_Reset.Execute';
        AxisData.Diag.tStepPreset := T#1S;

        xPowerRequest := FALSE;
        xResetExecute := FALSE;

        IF NOT fbReset.Busy THEN
            AxisData.Diag.iStep := E_AXIS_STATE.RESET_FINISH;
        END_IF;

    // --------------------------------------------------
    E_AXIS_STATE.RESET_FINISH:
    // --------------------------------------------------
        AxisData.Diag.sStepName := 'RESET_FINISH';
        AxisData.Diag.sWaitReason := 'Finishing reset';
        AxisData.Diag.tStepPreset := T#0S;

        xPowerRequest := FALSE;
        xResetExecute := FALSE;

        IF xDoResetAxis THEN
            AxisData.Error.dwAxisErrorLatched := DWORD#0;
        END_IF;
        IF xDoResetLogical THEN
            AxisData.Error.dwLogicalErrorLatched := DWORD#0;
            AxisData.Diag.xStepTimeout := FALSE;
        END_IF;

        xDoResetAxis := FALSE;
        xDoResetLogical := FALSE;

        // Финальная проверка
        IF AxisData.Error.dwAxisErrorActual <> DWORD#0 THEN
            AxisData.Diag.sWarningText := 'Axis error remains active after reset';
            uiResetWarningCode := WRN_RESET_AXIS_ACTIVE;
            AxisData.Error.dwAxisErrorLatched :=
                AxisData.Error.dwAxisErrorLatched OR AxisData.Error.dwAxisErrorActual;
            AxisData.Diag.iStep := E_AXIS_STATE.ERROR_RESET_MANAGER;

        ELSIF AxisData.Error.dwAxisErrorLatched <> DWORD#0 THEN
            AxisData.Diag.sWarningText := 'Latched axis error was not reset';
            uiResetWarningCode := WRN_RESET_AXIS_LATCHED;
            AxisData.Diag.iStep := E_AXIS_STATE.ERROR_RESET_MANAGER;

        ELSIF AxisData.Error.dwLogicalErrorLatched <> DWORD#0 THEN
            AxisData.Diag.sWarningText := 'Logical axis error was not reset';
            uiResetWarningCode := WRN_RESET_LOGICAL_ACTIVE;
            AxisData.Diag.iStep := E_AXIS_STATE.ERROR_RESET_MANAGER;

        ELSIF AxisData.Command.xGlobalError THEN
            AxisData.Diag.sWarningText := 'Global error is still active';
            uiResetWarningCode := WRN_RESET_GLOBAL_ERROR;
            AxisData.Diag.iStep := E_AXIS_STATE.ERROR_RESET_MANAGER;

        ELSE
            AxisData.Diag.iStep := E_AXIS_STATE.DISABLED;
        END_IF;

    // --------------------------------------------------
    ELSE  // неизвестное состояние
    // --------------------------------------------------
        AxisData.Error.dwLogicalErrorLatched :=
            AxisData.Error.dwLogicalErrorLatched OR LOG_UNKNOWN_STEP;
        AxisData.Diag.iLastErrorStep := TO_INT(AxisData.Diag.iStep);
        AxisData.Diag.iStep := E_AXIS_STATE.ERROR_RESET_MANAGER;

END_CASE;

// ======================================================
// 5. ТАЙМЕР ШАГА И КОНТРОЛЬ ТАЙМАУТА
// ======================================================
xStepChanged := (AxisData.Diag.iStep <> iPrevStep);
IF xStepChanged THEN
    iPrevStep := AxisData.Diag.iStep;
    xStepTimerEnable := FALSE;
ELSE
    xStepTimerEnable := TRUE;
END_IF;

tonStep(IN := xStepTimerEnable, PT := T#1000H);
AxisData.Diag.tStepElapsed := tonStep.ET;

tonStepTimeout(
    IN := xStepTimerEnable AND (AxisData.Diag.tStepPreset > T#0S),
    PT := AxisData.Diag.tStepPreset
);

IF tonStepTimeout.Q AND (AxisData.Diag.iStep <> E_AXIS_STATE.ERROR_RESET_MANAGER) THEN
    IF (AxisData.Diag.iStep = E_AXIS_STATE.RESET_AXIS_ERROR)
    OR (AxisData.Diag.iStep = E_AXIS_STATE.RESET_RELEASE) THEN
        AxisData.Diag.sWarningText := 'Axis reset timeout';
        uiResetWarningCode := WRN_RESET_TIMEOUT;
    END_IF;

    AxisData.Diag.xStepTimeout := TRUE;
    AxisData.Error.dwLogicalErrorLatched := AxisData.Error.dwLogicalErrorLatched OR LOG_STEP_TIMEOUT;
    AxisData.Diag.iLastErrorStep := TO_INT(AxisData.Diag.iStep);

    xResetExecute    := FALSE;
    xStopExecute     := FALSE;
    xHomeExecute     := FALSE;
    xMoveAbsExecute  := FALSE;
    xMoveRelExecute  := FALSE;
    xJogForwardExec  := FALSE;
    xJogBackwardExec := FALSE;

    AxisData.Diag.iStep := E_AXIS_STATE.ERROR_RESET_MANAGER;
END_IF;

IF uiResetWarningCode <> UINT#0 THEN
    AxisData.Diag.stWarning.uiCode := uiResetWarningCode;
    AxisData.Diag.stWarning.udiSequence := AxisData.Diag.stWarning.udiSequence + UDINT#1;
    IF AxisData.Diag.stWarning.udiSequence = UDINT#0 THEN
        AxisData.Diag.stWarning.udiSequence := UDINT#1;
    END_IF;
    xWarningPulse := TRUE;
END_IF;

// ======================================================
// 6. УДЕРЖАНИЕ ПРЕДУПРЕЖДЕНИЙ (TP)
// ======================================================
tpWarningHold(IN := xWarningPulse, PT := T#2S);
IF NOT tpWarningHold.Q THEN
    AxisData.Error.dwWarningLatched := DWORD#0;
    AxisData.Diag.sWarningText := '';
END_IF;
AxisData.Error.dwWarning := AxisData.Error.dwWarningLatched;
AxisData.Status.xWarning := (AxisData.Error.dwWarning <> DWORD#0);

// ======================================================
// 7. ВЫЗОВ MC-БЛОКОВ
// ======================================================
fbPower(
    Axis := Axis,
    // Enable активирует обработку MC_Power и не является командой питания.
    // Для штатного выключения FB продолжает выполняться, а силовые входы снимаются.
    Enable := TRUE,
    bRegulatorOn := xPowerRequest,
    bDriveStart := xPowerRequest
);

fbReset(
    Axis := Axis,
    Execute := xResetExecute
);

fbStop(
    Axis := Axis,
    Execute := xStopExecute,
    Deceleration := lrEffectiveDeceleration,
    Jerk := lrEffectiveJerk
);

fbJog(
    Axis := Axis,
    JogForward := xJogForwardExec,
    JogBackward := xJogBackwardExec,
    Velocity := lrEffectiveVelocity,
    Acceleration := lrEffectiveAcceleration,
    Deceleration := lrEffectiveDeceleration,
    Jerk := lrEffectiveJerk
);

fbHome(
    Axis := Axis,
    Execute := xHomeExecute,
    Position := AxisData.MotionParam.lrHomePosition
);

fbMoveAbsolute(
    Axis := Axis,
    Execute := xMoveAbsExecute,
    Position := AxisData.MotionParam.lrTargetPosition,
    Velocity := lrEffectiveVelocity,
    Acceleration := lrEffectiveAcceleration,
    Deceleration := lrEffectiveDeceleration,
    Jerk := lrEffectiveJerk,
    Direction := MC_DIRECTION.shortest,
    BufferMode := MC_BUFFER_MODE.Aborting
);

fbMoveRelative(
    Axis := Axis,
    Execute := xMoveRelExecute,
    Distance := AxisData.MotionParam.lrDistance,
    Velocity := lrEffectiveVelocity,
    Acceleration := lrEffectiveAcceleration,
    Deceleration := lrEffectiveDeceleration,
    Jerk := lrEffectiveJerk,
    BufferMode := MC_BUFFER_MODE.Aborting
);

fbReadPosition(
    Axis := Axis,
    Enable := TRUE
);

fbReadStatus(
    Axis := Axis,
    Enable := TRUE
);

fbReadAxisError(
    Axis := Axis,
    Enable := TRUE
);

// ======================================================
// 8. ИТОГОВЫЕ СТАТУСЫ (запись в структуру)
// ======================================================
AxisData.Status.xStandstill := fbReadStatus.Valid AND NOT AxisData.Status.xMotionBusy
	AND (fbReadStatus.StandStill OR fbReadStatus.Disabled OR fbReadStatus.Errorstop);
AxisData.Status.lrActualPosition := LREAL_TO_REAL(fbReadPosition.Position);

// Повторно собираем актуальные ошибки (для полноты)
AxisData.Error.dwAxisErrorActual := DWORD#0;
AxisData.Error.dwAxisErrorActual.0  := fbPower.Error;
AxisData.Error.dwAxisErrorActual.1  := fbReset.Error;
AxisData.Error.dwAxisErrorActual.2  := fbStop.Error;
AxisData.Error.dwAxisErrorActual.3  := fbJog.Error;
AxisData.Error.dwAxisErrorActual.4  := fbHome.Error;
AxisData.Error.dwAxisErrorActual.5  := fbMoveAbsolute.Error;
AxisData.Error.dwAxisErrorActual.6  := fbMoveRelative.Error;
AxisData.Error.dwAxisErrorActual.7  := fbReadPosition.Error;
AxisData.Error.dwAxisErrorActual.8  := fbReadStatus.Error;
AxisData.Error.dwAxisErrorActual.9  := fbReadStatus.Errorstop;
AxisData.Error.dwAxisErrorActual.10 := fbReadStatus.FBErrorOccured;
AxisData.Error.dwAxisErrorActual.11 := fbReadAxisError.AxisError;

xAxisErrorActual := (AxisData.Error.dwAxisErrorActual <> DWORD#0);

AxisData.Status.xLocalError :=
    fbPower.Error OR
    fbReset.Error OR
    fbStop.Error OR
    fbJog.Error OR
    fbHome.Error OR
    fbMoveAbsolute.Error OR
    fbMoveRelative.Error OR
    fbReadPosition.Error OR
    fbReadStatus.Error OR
    fbReadStatus.Errorstop OR
    fbReadStatus.FBErrorOccured OR
    fbReadAxisError.AxisError;

AxisData.Status.xMotionBusy :=
    fbStop.Busy OR
    fbJog.Busy OR
    fbHome.Busy OR
    fbMoveAbsolute.Busy OR
    fbMoveRelative.Busy;

xNeedMcReset :=
    fbReadStatus.Errorstop OR
    fbReadStatus.FBErrorOccured OR
    fbReadAxisError.AxisError;

AxisData.Error.dwAxisError := AxisData.Error.dwAxisErrorActual OR AxisData.Error.dwAxisErrorLatched;
AxisData.Error.dwLogicalError := AxisData.Error.dwLogicalErrorLatched;
AxisData.Error.dwAllError := AxisData.Error.dwAxisError OR AxisData.Error.dwLogicalError;
AxisData.Error.dwAlarmActive := AxisData.Error.dwAxisError
    OR SHL(AxisData.Error.dwLogicalError, 16);
AxisData.Error.dwDriveAxisErrorID := fbReadAxisError.AxisErrorID;

AxisData.Status.xAxisError := (AxisData.Error.dwAxisError <> DWORD#0);
AxisData.Status.xLogicalError := (AxisData.Error.dwLogicalError <> DWORD#0);
AxisData.Status.xAxisResetNeeded := AxisData.Status.xAxisError;
AxisData.Status.xLogicalResetNeeded := AxisData.Status.xLogicalError;

AxisData.Status.xError :=
    (AxisData.Diag.iStep = E_AXIS_STATE.ERROR_RESET_MANAGER) OR
    AxisData.Status.xAxisError OR
    AxisData.Status.xLogicalError OR
    AxisData.Command.xGlobalError;

AxisData.Status.xBusy :=
    fbPower.Busy OR
    fbReset.Busy OR
    AxisData.Status.xMotionBusy;

AxisData.Status.xCanStartMotion :=
    (AxisData.Diag.iStep = E_AXIS_STATE.READY) AND
    AxisData.Status.xPowered AND
    NOT AxisData.Status.xMotionBusy AND
    NOT AxisData.Status.xAxisError AND
    NOT AxisData.Status.xLogicalError AND
    NOT AxisData.Command.xGlobalError;

// ======================================================
// 9. ТЕКСТ ОШИБКИ И ID
// ======================================================
AxisData.Diag.sErrorText := '';
AxisData.Diag.udiActualErrorID := 0;

IF (AxisData.Error.dwLogicalError AND LOG_POWER_PERMIT_LOST) <> DWORD#0 THEN
    AxisData.Diag.sErrorText := 'Power permit lost';
    AxisData.Diag.udiActualErrorID := 1001;

ELSIF (AxisData.Error.dwLogicalError AND LOG_GLOBAL_DURING_POWER) <> DWORD#0 THEN
    AxisData.Diag.sErrorText := 'Global error during power on';
    AxisData.Diag.udiActualErrorID := 1002;

ELSIF (AxisData.Error.dwLogicalError AND LOG_GLOBAL_DURING_READY) <> DWORD#0 THEN
    AxisData.Diag.sErrorText := 'Global error in READY state';
    AxisData.Diag.udiActualErrorID := 2000;

ELSIF (AxisData.Error.dwLogicalError AND LOG_GLOBAL_DURING_MOTION) <> DWORD#0 THEN
    AxisData.Diag.sErrorText := 'Global error during motion';
    AxisData.Diag.udiActualErrorID := 2100;

ELSIF (AxisData.Error.dwLogicalError AND LOG_JOG_CONFLICT) <> DWORD#0 THEN
    AxisData.Diag.sErrorText := 'Jog positive and negative active together';
    AxisData.Diag.udiActualErrorID := 2001;

ELSIF (AxisData.Error.dwLogicalError AND LOG_MOVE_ABS_NOT_HOMED) <> DWORD#0 THEN
    AxisData.Diag.sErrorText := 'MoveAbsolute denied: axis not homed';
    AxisData.Diag.udiActualErrorID := 1200;

ELSIF (AxisData.Error.dwLogicalError AND LOG_MOVE_REL_NOT_HOMED) <> DWORD#0 THEN
    AxisData.Diag.sErrorText := 'MoveRelative denied: axis not homed';
    AxisData.Diag.udiActualErrorID := 1300;

ELSIF (AxisData.Error.dwLogicalError AND LOG_STEP_TIMEOUT) <> DWORD#0 THEN
    AxisData.Diag.sErrorText := 'Step timeout';
    AxisData.Diag.udiActualErrorID := 9000 + INT_TO_UDINT(AxisData.Diag.iLastErrorStep);

ELSIF (AxisData.Error.dwLogicalError AND LOG_UNKNOWN_STEP) <> DWORD#0 THEN
    AxisData.Diag.sErrorText := 'Unknown axis step';
    AxisData.Diag.udiActualErrorID := 9999;

ELSIF (AxisData.Error.dwAxisError AND AXE_MC_POWER_ERROR) <> DWORD#0 THEN
    AxisData.Diag.sErrorText := 'MC_Power error';
    AxisData.Diag.udiActualErrorID := TO_UDINT(fbPower.ErrorID);

ELSIF (AxisData.Error.dwAxisError AND AXE_MC_RESET_ERROR) <> DWORD#0 THEN
    AxisData.Diag.sErrorText := 'MC_Reset error';
    AxisData.Diag.udiActualErrorID := TO_UDINT(fbReset.ErrorID);

ELSIF (AxisData.Error.dwAxisError AND AXE_MC_STOP_ERROR) <> DWORD#0 THEN
    AxisData.Diag.sErrorText := 'MC_Stop error';
    AxisData.Diag.udiActualErrorID := TO_UDINT(fbStop.ErrorID);

ELSIF (AxisData.Error.dwAxisError AND AXE_MC_JOG_ERROR) <> DWORD#0 THEN
    AxisData.Diag.sErrorText := 'MC_Jog error';
    AxisData.Diag.udiActualErrorID := TO_UDINT(fbJog.ErrorID);

ELSIF (AxisData.Error.dwAxisError AND AXE_MC_HOME_ERROR) <> DWORD#0 THEN
    AxisData.Diag.sErrorText := 'MC_Home error';
    AxisData.Diag.udiActualErrorID := TO_UDINT(fbHome.ErrorID);

ELSIF (AxisData.Error.dwAxisError AND AXE_MC_MOVE_ABS_ERROR) <> DWORD#0 THEN
    AxisData.Diag.sErrorText := 'MC_MoveAbsolute error';
    AxisData.Diag.udiActualErrorID := TO_UDINT(fbMoveAbsolute.ErrorID);

ELSIF (AxisData.Error.dwAxisError AND AXE_MC_MOVE_REL_ERROR) <> DWORD#0 THEN
    AxisData.Diag.sErrorText := 'MC_MoveRelative error';
    AxisData.Diag.udiActualErrorID := TO_UDINT(fbMoveRelative.ErrorID);

ELSIF (AxisData.Error.dwAxisError AND AXE_READ_POS_ERROR) <> DWORD#0 THEN
    AxisData.Diag.sErrorText := 'MC_ReadActualPosition error';
    AxisData.Diag.udiActualErrorID := TO_UDINT(fbReadPosition.ErrorID);

ELSIF (AxisData.Error.dwAxisError AND AXE_READ_STATUS_ERROR) <> DWORD#0 THEN
    AxisData.Diag.sErrorText := 'MC_ReadStatus error';
    AxisData.Diag.udiActualErrorID := TO_UDINT(fbReadStatus.ErrorID);

ELSIF (AxisData.Error.dwAxisError AND AXE_ERRORSTOP) <> DWORD#0 THEN
    AxisData.Diag.sErrorText := 'Axis Errorstop active';
    AxisData.Diag.udiActualErrorID := 3001;

ELSIF (AxisData.Error.dwAxisError AND AXE_FB_ERROR_OCCURRED) <> DWORD#0 THEN
    AxisData.Diag.sErrorText := 'SoftMotion FBErrorOccured active';
    AxisData.Diag.udiActualErrorID := 3002;

ELSIF (AxisData.Error.dwAxisError AND AXE_COMMAND_ABORTED) <> DWORD#0 THEN
    AxisData.Diag.sErrorText := 'Motion command aborted';
    AxisData.Diag.udiActualErrorID := 3003;

ELSIF (AxisData.Error.dwAxisError AND AXE_UNKNOWN_ACTUAL_ERROR) <> DWORD#0 THEN
    AxisData.Diag.sErrorText := 'Unknown actual axis error';
    AxisData.Diag.udiActualErrorID := 3004;

ELSIF (AxisData.Error.dwAxisError AND AXE_DRIVE_AXIS_ERROR) <> DWORD#0 THEN
    AxisData.Diag.sErrorText := 'Drive axis error active';
    AxisData.Diag.udiActualErrorID := DWORD_TO_UDINT(fbReadAxisError.AxisErrorID);

ELSIF (AxisData.Error.dwAxisError AND AXE_POWER_FEEDBACK_LOST) <> DWORD#0 THEN
    AxisData.Diag.sErrorText := 'Drive power feedback lost';
    AxisData.Diag.udiActualErrorID := 3005;

ELSIF AxisData.Command.xGlobalError THEN
    AxisData.Diag.sErrorText := 'Global error active';
    AxisData.Diag.udiActualErrorID := 5000;
END_IF;

IF AxisData.Diag.udiActualErrorID <> 0 THEN
    AxisData.Diag.udiLastErrorID := AxisData.Diag.udiActualErrorID;
END_IF;

// Сохраняем последнюю ненулевую ошибку и формируем удобное представление для HMI.
IF (AxisData.Error.dwAxisError <> DWORD#0)
OR (AxisData.Error.dwLogicalError <> DWORD#0) THEN
	AxisData.Error.dwAxisErrorLast := AxisData.Error.dwAxisError;
	AxisData.Error.dwLogicalErrorLast := AxisData.Error.dwLogicalError;
END_IF;

AxisData.Error.stErrorActive := UpdateErrorView(
	dwAxisError := AxisData.Error.dwAxisError,
	dwLogicalError := AxisData.Error.dwLogicalError
);
AxisData.Error.stErrorLast := UpdateErrorView(
    dwAxisError := AxisData.Error.dwAxisErrorLast,
    dwLogicalError := AxisData.Error.dwLogicalErrorLast
);

FaultStatus.xResetAllowed := AxisData.Status.xError
	AND xResetPermit
	AND NOT AxisData.Command.xGlobalError
	AND NOT FaultStatus.xBusy;

METHOD UpdateErrorView : ST_AXIS_ERROR
VAR_INPUT
	dwAxisError   : DWORD; // Маска ошибок SoftMotion и привода
	dwLogicalError: DWORD; // Маска логических ошибок оси
END_VAR
VAR
	stError : ST_AXIS_ERROR; // Представление ошибок отдельными флагами
END_VAR
stError.MC_POWER_ERROR := (dwAxisError AND AXE_MC_POWER_ERROR) <> DWORD#0;
stError.MC_RESET_ERROR := (dwAxisError AND AXE_MC_RESET_ERROR) <> DWORD#0;
stError.MC_STOP_ERROR := (dwAxisError AND AXE_MC_STOP_ERROR) <> DWORD#0;
stError.MC_JOG_ERROR := (dwAxisError AND AXE_MC_JOG_ERROR) <> DWORD#0;
stError.MC_HOME_ERROR := (dwAxisError AND AXE_MC_HOME_ERROR) <> DWORD#0;
stError.MC_MOVE_ABS_ERROR := (dwAxisError AND AXE_MC_MOVE_ABS_ERROR) <> DWORD#0;
stError.MC_MOVE_REL_ERROR := (dwAxisError AND AXE_MC_MOVE_REL_ERROR) <> DWORD#0;
stError.READ_POSITION_ERROR := (dwAxisError AND AXE_READ_POS_ERROR) <> DWORD#0;
stError.READ_STATUS_ERROR := (dwAxisError AND AXE_READ_STATUS_ERROR) <> DWORD#0;
stError.AXIS_ERRORSTOP := (dwAxisError AND AXE_ERRORSTOP) <> DWORD#0;
stError.FB_ERROR_OCCURRED := (dwAxisError AND AXE_FB_ERROR_OCCURRED) <> DWORD#0;
stError.COMMAND_ABORTED := (dwAxisError AND AXE_COMMAND_ABORTED) <> DWORD#0;
stError.UNKNOWN_AXIS_ERROR := (dwAxisError AND AXE_UNKNOWN_ACTUAL_ERROR) <> DWORD#0;
stError.DRIVE_AXIS_ERROR := (dwAxisError AND AXE_DRIVE_AXIS_ERROR) <> DWORD#0;
stError.POWER_FEEDBACK_LOST := (dwAxisError AND AXE_POWER_FEEDBACK_LOST) <> DWORD#0;

stError.POWER_PERMIT_LOST := (dwLogicalError AND LOG_POWER_PERMIT_LOST) <> DWORD#0;
stError.GLOBAL_DURING_POWER := (dwLogicalError AND LOG_GLOBAL_DURING_POWER) <> DWORD#0;
stError.GLOBAL_DURING_READY := (dwLogicalError AND LOG_GLOBAL_DURING_READY) <> DWORD#0;
stError.GLOBAL_DURING_MOTION := (dwLogicalError AND LOG_GLOBAL_DURING_MOTION) <> DWORD#0;
stError.JOG_CONFLICT := (dwLogicalError AND LOG_JOG_CONFLICT) <> DWORD#0;
stError.MOVE_ABS_NOT_HOMED := (dwLogicalError AND LOG_MOVE_ABS_NOT_HOMED) <> DWORD#0;
stError.MOVE_REL_NOT_HOMED := (dwLogicalError AND LOG_MOVE_REL_NOT_HOMED) <> DWORD#0;
stError.STEP_TIMEOUT := (dwLogicalError AND LOG_STEP_TIMEOUT) <> DWORD#0;
stError.UNKNOWN_STEP := (dwLogicalError AND LOG_UNKNOWN_STEP) <> DWORD#0;

UpdateErrorView := stError;
END_METHOD

END_FUNCTION_BLOCK

// Device/Application/FB/FB_FAULT_INJECTOR/FB_AXIS_FAULT_INJECTOR
FUNCTION_BLOCK FB_AXIS_FAULT_INJECTOR
VAR_INPUT
	Request      : ST_AXIS_FAULT_REQUEST; // Запрос тестовой логической ошибки оси
	xOwnerAllowed: BOOL; // Безопасные условия, рассчитанные FB_AXIS
END_VAR
VAR_OUTPUT
	xJogConflict : BOOL; // Одноцикловая пара Jog+ и Jog- для штатной проверки
	Status       : ST_FAULT_INJECTION_STATUS; // Состояние источника для HMI
END_VAR
VAR
	rtJogConflict : R_TRIG; // Фронт команды HMI
END_VAR

rtJogConflict(CLK := Request.xJogConflict);

xJogConflict := FALSE;
Status.xRejected := FALSE;
Status.xAllowed := Request.xEnabled AND xOwnerAllowed;
Status.xBusy := FALSE;
Status.xResetAllowed := FALSE;

IF rtJogConflict.Q THEN
	IF Status.xAllowed THEN
		xJogConflict := TRUE;
	ELSE
		Status.xRejected := TRUE;
		Status.udiRejectSequence := Status.udiRejectSequence + UDINT#1;
		IF Status.udiRejectSequence = UDINT#0 THEN
			Status.udiRejectSequence := UDINT#1;
		END_IF;
	END_IF;
END_IF;

Status.xActive := xJogConflict;

END_FUNCTION_BLOCK

// Device/Application/FB/FB_AXIS_GROUP
FUNCTION_BLOCK FB_AXIS_GROUP
VAR_INPUT
	FaultRequest : ST_AXIS_GROUP_FAULT_REQUEST; // Единый контракт диагностической инъекции
	xResetPermit : BOOL; // Общий сброс разрешён ручным режимом и остановленной ячейкой
	xAxesPowered : BOOL; // Питанием физических осей владеют FB_AXIS; группа только наблюдает готовность
	lrVelocityOverride : LREAL; // Live override скорости групповых движений, 0.001..1.0
END_VAR
VAR_OUTPUT
	FaultStatus : ST_FAULT_INJECTION_STATUS; // Состояние инжектора для HMI
END_VAR
VAR
	// Внутренние исполняемые булевые переменные
	xEnable      : BOOL; // Импульс включения группы
	xDisable     : BOOL; // Импульс отключения группы
	xReset       : BOOL; // Импульс сброса ошибок
	xResetMC     : BOOL; // Выполняется сброс SoftMotion
	xMoveDirect  : BOOL; // Выполняется прямое перемещение
	xMoveLinear  : BOOL; // Выполняется линейное перемещение
	xStopCmd     : BOOL; // Выполняется остановка
	xHaltCmd     : BOOL; // Выполняется плавная остановка
	lrAppliedVelocityOverride : LREAL; // Коэффициент после защитного ограничения PLC
	xVelocityOverrideEnable : BOOL; // Запись live override разрешена только в рабочих состояниях без MC_GroupStop
	xFaultAllowed : BOOL; // Безопасные условия тестового запуска
	
	iPrevStep : E_AXIS_GROUP_STATE; // Предыдущий шаг автомата
	
